(* IEC 61131-3 sources: plc-st-coding-agent/progress/evidence/f14_v11_public_20261113/jobs/custom_deepseek-v4pro, 104 files *)

(* ---- public-easy-01.candidate_01.st ---- *)
(* ENGINEERING_CONTRACT
Outputs by state (state is persistent across scans):
- Pump_Motor: ON in CLEANING; starts when bottleSensor TRUE from IDLE; OFF on cleaningConfirmButton. Retained while CLEANING, even if bottleSensor falls (PUB001/PUB002).
- Filling_Valve: ON in FILLING; starts on cleaningConfirmButton in CLEANING; OFF on fillingConfirmButton (PUB002/PUB003).
- Capping_Machine: ON in CAPPING; starts on fillingConfirmButton in FILLING; OFF on cappingConfirmButton (PUB003/PUB004).
- Packing_Machine: ON in PACKING; starts on cappingConfirmButton in CAPPING; OFF on packingConfirmButton (PUB004/PUB005).
- Completion_Light: ON in COMPLETE; starts on packingConfirmButton in PACKING; reset by finishedButton (PUB005/PUB006/PUB007).
Same-scan priority: one state transition per call via ELSIF chain; outputs are assigned after transition using final state.
Buttons are treated as level-sensitive; pulse width/protocol unspecified.
*)
(* CONTRACT_RULES [] *)

FUNCTION_BLOCK FillingLineControl
VAR_INPUT
    bottleSensor: BOOL;
    cleaningConfirmButton: BOOL;
    fillingConfirmButton: BOOL;
    cappingConfirmButton: BOOL;
    packingConfirmButton: BOOL;
    finishedButton: BOOL;
END_VAR
VAR_OUTPUT
    Pump_Motor: BOOL;
    Filling_Valve: BOOL;
    Capping_Machine: BOOL;
    Packing_Machine: BOOL;
    Completion_Light: BOOL;
END_VAR
VAR
    step: INT := 0; (* 0=IDLE, 1=CLEANING, 2=FILLING, 3=CAPPING, 4=PACKING, 5=COMPLETE *)
END_VAR

(* State transitions: at most one per scan *)
IF step = 0 THEN
    IF bottleSensor THEN
        step := 1;
    END_IF;
ELSIF step = 1 THEN
    IF cleaningConfirmButton THEN
        step := 2;
    END_IF;
ELSIF step = 2 THEN
    IF fillingConfirmButton THEN
        step := 3;
    END_IF;
ELSIF step = 3 THEN
    IF cappingConfirmButton THEN
        step := 4;
    END_IF;
ELSIF step = 4 THEN
    IF packingConfirmButton THEN
        step := 5;
    END_IF;
ELSIF step = 5 THEN
    IF finishedButton THEN
        step := 0;
    END_IF;
END_IF;

(* Output mapping based on final state *)
CASE step OF
    0:
        Pump_Motor := FALSE;
        Filling_Valve := FALSE;
        Capping_Machine := FALSE;
        Packing_Machine := FALSE;
        Completion_Light := FALSE;

    1:
        Pump_Motor := TRUE;
        Filling_Valve := FALSE;
        Capping_Machine := FALSE;
        Packing_Machine := FALSE;
        Completion_Light := FALSE;

    2:
        Pump_Motor := FALSE;
        Filling_Valve := TRUE;
        Capping_Machine := FALSE;
        Packing_Machine := FALSE;
        Completion_Light := FALSE;

    3:
        Pump_Motor := FALSE;
        Filling_Valve := FALSE;
        Capping_Machine := TRUE;
        Packing_Machine := FALSE;
        Completion_Light := FALSE;

    4:
        Pump_Motor := FALSE;
        Filling_Valve := FALSE;
        Capping_Machine := FALSE;
        Packing_Machine := TRUE;
        Completion_Light := FALSE;

    5:
        Pump_Motor := FALSE;
        Filling_Valve := FALSE;
        Capping_Machine := FALSE;
        Packing_Machine := FALSE;
        Completion_Light := TRUE;

    ELSE
        Pump_Motor := FALSE;
        Filling_Valve := FALSE;
        Capping_Machine := FALSE;
        Packing_Machine := FALSE;
        Completion_Light := FALSE;
END_CASE;

(* ---- public-easy-01.candidate_02.st ---- *)
(* ENGINEERING_CONTRACT
Outputs by state (state is persistent across scans):
- Pump_Motor: ON in CLEANING; starts when bottleSensor TRUE from IDLE; OFF on cleaningConfirmButton. Retained while CLEANING, even if bottleSensor falls (PUB001/PUB002).
- Filling_Valve: ON in FILLING; starts on cleaningConfirmButton in CLEANING; OFF on fillingConfirmButton (PUB002/PUB003).
- Capping_Machine: ON in CAPPING; starts on fillingConfirmButton in FILLING; OFF on cappingConfirmButton (PUB003/PUB004).
- Packing_Machine: ON in PACKING; starts on cappingConfirmButton in CAPPING; OFF on packingConfirmButton (PUB004/PUB005).
- Completion_Light: ON in COMPLETE; starts on packingConfirmButton in PACKING; reset by finishedButton (PUB005/PUB006/PUB007).
Same-scan priority: one state transition per call via ELSIF chain; outputs are assigned after transition using final state.
Buttons are treated as level-sensitive; pulse width/protocol unspecified.
*)
(* CONTRACT_RULES [] *)

FUNCTION_BLOCK FillingLineControl
VAR_INPUT
    bottleSensor: BOOL;
    cleaningConfirmButton: BOOL;
    fillingConfirmButton: BOOL;
    cappingConfirmButton: BOOL;
    packingConfirmButton: BOOL;
    finishedButton: BOOL;
END_VAR
VAR_OUTPUT
    Pump_Motor: BOOL;
    Filling_Valve: BOOL;
    Capping_Machine: BOOL;
    Packing_Machine: BOOL;
    Completion_Light: BOOL;
END_VAR
VAR
    step: INT := 0; (* 0=IDLE, 1=CLEANING, 2=FILLING, 3=CAPPING, 4=PACKING, 5=COMPLETE *)
END_VAR

(* State transitions: at most one per scan *)
IF step = 0 THEN
    IF bottleSensor THEN
        step := 1;
    END_IF;
ELSIF step = 1 THEN
    IF cleaningConfirmButton THEN
        step := 2;
    END_IF;
ELSIF step = 2 THEN
    IF fillingConfirmButton THEN
        step := 3;
    END_IF;
ELSIF step = 3 THEN
    IF cappingConfirmButton THEN
        step := 4;
    END_IF;
ELSIF step = 4 THEN
    IF packingConfirmButton THEN
        step := 5;
    END_IF;
ELSIF step = 5 THEN
    IF finishedButton THEN
        step := 0;
    END_IF;
END_IF;

(* Output mapping based on final state *)
CASE step OF
    0:
        Pump_Motor := FALSE;
        Filling_Valve := FALSE;
        Capping_Machine := FALSE;
        Packing_Machine := FALSE;
        Completion_Light := FALSE;

    1:
        Pump_Motor := TRUE;
        Filling_Valve := FALSE;
        Capping_Machine := FALSE;
        Packing_Machine := FALSE;
        Completion_Light := FALSE;

    2:
        Pump_Motor := FALSE;
        Filling_Valve := TRUE;
        Capping_Machine := FALSE;
        Packing_Machine := FALSE;
        Completion_Light := FALSE;

    3:
        Pump_Motor := FALSE;
        Filling_Valve := FALSE;
        Capping_Machine := TRUE;
        Packing_Machine := FALSE;
        Completion_Light := FALSE;

    4:
        Pump_Motor := FALSE;
        Filling_Valve := FALSE;
        Capping_Machine := FALSE;
        Packing_Machine := TRUE;
        Completion_Light := FALSE;

    5:
        Pump_Motor := FALSE;
        Filling_Valve := FALSE;
        Capping_Machine := FALSE;
        Packing_Machine := FALSE;
        Completion_Light := TRUE;

    ELSE
        Pump_Motor := FALSE;
        Filling_Valve := FALSE;
        Capping_Machine := FALSE;
        Packing_Machine := FALSE;
        Completion_Light := FALSE;
END_CASE;

END_FUNCTION_BLOCK

(* ---- public-easy-01.candidate_03.st ---- *)
(* ENGINEERING_CONTRACT
Outputs by state (state is persistent across scans):
- Pump_Motor: ON in CLEANING; starts when bottleSensor TRUE from IDLE; OFF on cleaningConfirmButton. Retained while CLEANING, even if bottleSensor falls (PUB001/PUB002).
- Filling_Valve: ON in FILLING; starts on cleaningConfirmButton in CLEANING; OFF on fillingConfirmButton (PUB002/PUB003).
- Capping_Machine: ON in CAPPING; starts on fillingConfirmButton in FILLING; OFF on cappingConfirmButton (PUB003/PUB004).
- Packing_Machine: ON in PACKING; starts on cappingConfirmButton in CAPPING; OFF on packingConfirmButton (PUB004/PUB005).
- Completion_Light: ON in COMPLETE; starts on packingConfirmButton in PACKING; reset by finishedButton (PUB005/PUB006/PUB007).
Same-scan priority:
- Primary ELSIF chain processes one normal step.
- If finishedButton resets to IDLE and bottleSensor is already TRUE, re-enter CLEANING immediately in same scan.
Outputs are assigned after transition logic using final state.
Buttons are treated as level-sensitive; pulse width/protocol unspecified.
*)
(* CONTRACT_RULES [] *)

FUNCTION_BLOCK FillingLineControl
VAR_INPUT
    bottleSensor: BOOL;
    cleaningConfirmButton: BOOL;
    fillingConfirmButton: BOOL;
    cappingConfirmButton: BOOL;
    packingConfirmButton: BOOL;
    finishedButton: BOOL;
END_VAR
VAR_OUTPUT
    Pump_Motor: BOOL;
    Filling_Valve: BOOL;
    Capping_Machine: BOOL;
    Packing_Machine: BOOL;
    Completion_Light: BOOL;
END_VAR
VAR
    step: INT := 0; (* 0=IDLE, 1=CLEANING, 2=FILLING, 3=CAPPING, 4=PACKING, 5=COMPLETE *)
END_VAR

(* Primary state transitions: at most one normal step per scan *)
IF step = 0 THEN
    IF bottleSensor THEN
        step := 1;
    END_IF;
ELSIF step = 1 THEN
    IF cleaningConfirmButton THEN
        step := 2;
    END_IF;
ELSIF step = 2 THEN
    IF fillingConfirmButton THEN
        step := 3;
    END_IF;
ELSIF step = 3 THEN
    IF cappingConfirmButton THEN
        step := 4;
    END_IF;
ELSIF step = 4 THEN
    IF packingConfirmButton THEN
        step := 5;
    END_IF;
ELSIF step = 5 THEN
    IF finishedButton THEN
        step := 0;
    END_IF;
END_IF;

(* Same-scan reactivation: if finished just reset state to IDLE and a bottle is
   already detected, start cleaning immediately instead of waiting one scan. *)
IF step = 0 THEN
    IF bottleSensor THEN
        step := 1;
    END_IF;
END_IF;

(* Output mapping based on final state *)
CASE step OF
    0:
        Pump_Motor := FALSE;
        Filling_Valve := FALSE;
        Capping_Machine := FALSE;
        Packing_Machine := FALSE;
        Completion_Light := FALSE;

    1:
        Pump_Motor := TRUE;
        Filling_Valve := FALSE;
        Capping_Machine := FALSE;
        Packing_Machine := FALSE;
        Completion_Light := FALSE;

    2:
        Pump_Motor := FALSE;
        Filling_Valve := TRUE;
        Capping_Machine := FALSE;
        Packing_Machine := FALSE;
        Completion_Light := FALSE;

    3:
        Pump_Motor := FALSE;
        Filling_Valve := FALSE;
        Capping_Machine := TRUE;
        Packing_Machine := FALSE;
        Completion_Light := FALSE;

    4:
        Pump_Motor := FALSE;
        Filling_Valve := FALSE;
        Capping_Machine := FALSE;
        Packing_Machine := TRUE;
        Completion_Light := FALSE;

    5:
        Pump_Motor := FALSE;
        Filling_Valve := FALSE;
        Capping_Machine := FALSE;
        Packing_Machine := FALSE;
        Completion_Light := TRUE;

    ELSE
        Pump_Motor := FALSE;
        Filling_Valve := FALSE;
        Capping_Machine := FALSE;
        Packing_Machine := FALSE;
        Completion_Light := FALSE;
END_CASE;

END_FUNCTION_BLOCK

(* ---- public-easy-01.candidate_04.st ---- *)
(* ENGINEERING_CONTRACT
Outputs by state (state is persistent across scans):
- Pump_Motor: ON in CLEANING; starts when bottleSensor TRUE from IDLE; OFF on cleaningConfirmButton. Retained while CLEANING, even if bottleSensor falls (PUB001/PUB002).
- Filling_Valve: ON in FILLING; starts on cleaningConfirmButton in CLEANING; OFF on fillingConfirmButton (PUB002/PUB003).
- Capping_Machine: ON in CAPPING; starts on fillingConfirmButton in FILLING; OFF on cappingConfirmButton (PUB003/PUB004).
- Packing_Machine: ON in PACKING; starts on cappingConfirmButton in CAPPING; OFF on packingConfirmButton (PUB004/PUB005).
- Completion_Light: ON in COMPLETE; starts on packingConfirmButton in PACKING; reset by finishedButton (PUB005/PUB006/PUB007).
Same-scan priority:
- Primary ELSIF chain processes one normal step.
- If finishedButton resets to IDLE and bottleSensor is already TRUE, re-enter CLEANING immediately in same scan.
Outputs are assigned after transition logic using final state.
Buttons are treated as level-sensitive; pulse width/protocol unspecified.
*)
(* CONTRACT_RULES [
  {"kind":"hold_until_reset","output":"Pump_Motor","set_input":"bottleSensor","reset_input":"cleaningConfirmButton"},
  {"kind":"hold_until_reset","output":"Filling_Valve","set_input":"cleaningConfirmButton","reset_input":"fillingConfirmButton"},
  {"kind":"hold_until_reset","output":"Capping_Machine","set_input":"fillingConfirmButton","reset_input":"cappingConfirmButton"},
  {"kind":"hold_until_reset","output":"Packing_Machine","set_input":"cappingConfirmButton","reset_input":"packingConfirmButton"},
  {"kind":"hold_until_reset","output":"Completion_Light","set_input":"packingConfirmButton","reset_input":"finishedButton"}
] *)

FUNCTION_BLOCK FillingLineControl
VAR_INPUT
    bottleSensor: BOOL;
    cleaningConfirmButton: BOOL;
    fillingConfirmButton: BOOL;
    cappingConfirmButton: BOOL;
    packingConfirmButton: BOOL;
    finishedButton: BOOL;
END_VAR
VAR_OUTPUT
    Pump_Motor: BOOL;
    Filling_Valve: BOOL;
    Capping_Machine: BOOL;
    Packing_Machine: BOOL;
    Completion_Light: BOOL;
END_VAR
VAR
    step: INT := 0; (* 0=IDLE, 1=CLEANING, 2=FILLING, 3=CAPPING, 4=PACKING, 5=COMPLETE *)
END_VAR

(* Primary state transitions: at most one normal step per scan *)
IF step = 0 THEN
    IF bottleSensor THEN
        step := 1;
    END_IF;
ELSIF step = 1 THEN
    IF cleaningConfirmButton THEN
        step := 2;
    END_IF;
ELSIF step = 2 THEN
    IF fillingConfirmButton THEN
        step := 3;
    END_IF;
ELSIF step = 3 THEN
    IF cappingConfirmButton THEN
        step := 4;
    END_IF;
ELSIF step = 4 THEN
    IF packingConfirmButton THEN
        step := 5;
    END_IF;
ELSIF step = 5 THEN
    IF finishedButton THEN
        step := 0;
    END_IF;
END_IF;

(* Same-scan reactivation: if finished just reset state to IDLE and a bottle is
   already detected, start cleaning immediately instead of waiting one scan. *)
IF step = 0 THEN
    IF bottleSensor THEN
        step := 1;
    END_IF;
END_IF;

(* Output mapping based on final state *)
CASE step OF
    0:
        Pump_Motor := FALSE;
        Filling_Valve := FALSE;
        Capping_Machine := FALSE;
        Packing_Machine := FALSE;
        Completion_Light := FALSE;

    1:
        Pump_Motor := TRUE;
        Filling_Valve := FALSE;
        Capping_Machine := FALSE;
        Packing_Machine := FALSE;
        Completion_Light := FALSE;

    2:
        Pump_Motor := FALSE;
        Filling_Valve := TRUE;
        Capping_Machine := FALSE;
        Packing_Machine := FALSE;
        Completion_Light := FALSE;

    3:
        Pump_Motor := FALSE;
        Filling_Valve := FALSE;
        Capping_Machine := TRUE;
        Packing_Machine := FALSE;
        Completion_Light := FALSE;

    4:
        Pump_Motor := FALSE;
        Filling_Valve := FALSE;
        Capping_Machine := FALSE;
        Packing_Machine := TRUE;
        Completion_Light := FALSE;

    5:
        Pump_Motor := FALSE;
        Filling_Valve := FALSE;
        Capping_Machine := FALSE;
        Packing_Machine := FALSE;
        Completion_Light := TRUE;

    ELSE
        Pump_Motor := FALSE;
        Filling_Valve := FALSE;
        Capping_Machine := FALSE;
        Packing_Machine := FALSE;
        Completion_Light := FALSE;
END_CASE;

END_FUNCTION_BLOCK

(* ---- public-easy-01.raw_candidate_01.st ---- *)
(* ENGINEERING_CONTRACT
Outputs by state (state is persistent across scans):
- Pump_Motor: ON in CLEANING; starts when bottleSensor TRUE from IDLE; OFF on cleaningConfirmButton. Retained while CLEANING, even if bottleSensor falls (PUB001/PUB002).
- Filling_Valve: ON in FILLING; starts on cleaningConfirmButton in CLEANING; OFF on fillingConfirmButton (PUB002/PUB003).
- Capping_Machine: ON in CAPPING; starts on fillingConfirmButton in FILLING; OFF on cappingConfirmButton (PUB003/PUB004).
- Packing_Machine: ON in PACKING; starts on cappingConfirmButton in CAPPING; OFF on packingConfirmButton (PUB004/PUB005).
- Completion_Light: ON in COMPLETE; starts on packingConfirmButton in PACKING; reset by finishedButton (PUB005/PUB006/PUB007).
Same-scan priority: one state transition per call via ELSIF chain; outputs are assigned after transition using final state.
Buttons are treated as level-sensitive; pulse width/protocol unspecified.
*)
(* CONTRACT_RULES [] *)

FUNCTION_BLOCK FillingLineControl
VAR_INPUT
    bottleSensor: BOOL;
    cleaningConfirmButton: BOOL;
    fillingConfirmButton: BOOL;
    cappingConfirmButton: BOOL;
    packingConfirmButton: BOOL;
    finishedButton: BOOL;
END_VAR
VAR_OUTPUT
    Pump_Motor: BOOL;
    Filling_Valve: BOOL;
    Capping_Machine: BOOL;
    Packing_Machine: BOOL;
    Completion_Light: BOOL;
END_VAR
VAR
    step: INT := 0; (* 0=IDLE, 1=CLEANING, 2=FILLING, 3=CAPPING, 4=PACKING, 5=COMPLETE *)
END_VAR

(* State transitions: at most one per scan *)
IF step = 0 THEN
    IF bottleSensor THEN
        step := 1;
    END_IF;
ELSIF step = 1 THEN
    IF cleaningConfirmButton THEN
        step := 2;
    END_IF;
ELSIF step = 2 THEN
    IF fillingConfirmButton THEN
        step := 3;
    END_IF;
ELSIF step = 3 THEN
    IF cappingConfirmButton THEN
        step := 4;
    END_IF;
ELSIF step = 4 THEN
    IF packingConfirmButton THEN
        step := 5;
    END_IF;
ELSIF step = 5 THEN
    IF finishedButton THEN
        step := 0;
    END_IF;
END_IF;

(* Output mapping based on final state *)
CASE step OF
    0:
        Pump_Motor := FALSE;
        Filling_Valve := FALSE;
        Capping_Machine := FALSE;
        Packing_Machine := FALSE;
        Completion_Light := FALSE;

    1:
        Pump_Motor := TRUE;
        Filling_Valve := FALSE;
        Capping_Machine := FALSE;
        Packing_Machine := FALSE;
        Completion_Light := FALSE;

    2:
        Pump_Motor := FALSE;
        Filling_Valve := TRUE;
        Capping_Machine := FALSE;
        Packing_Machine := FALSE;
        Completion_Light := FALSE;

    3:
        Pump_Motor := FALSE;
        Filling_Valve := FALSE;
        Capping_Machine := TRUE;
        Packing_Machine := FALSE;
        Completion_Light := FALSE;

    4:
        Pump_Motor := FALSE;
        Filling_Valve := FALSE;
        Capping_Machine := FALSE;
        Packing_Machine := TRUE;
        Completion_Light := FALSE;

    5:
        Pump_Motor := FALSE;
        Filling_Valve := FALSE;
        Capping_Machine := FALSE;
        Packing_Machine := FALSE;
        Completion_Light := TRUE;

    ELSE
        Pump_Motor := FALSE;
        Filling_Valve := FALSE;
        Capping_Machine := FALSE;
        Packing_Machine := FALSE;
        Completion_Light := FALSE;
END_CASE;

(* ---- public-easy-01.raw_candidate_02.st ---- *)
(* ENGINEERING_CONTRACT
Outputs by state (state is persistent across scans):
- Pump_Motor: ON in CLEANING; starts when bottleSensor TRUE from IDLE; OFF on cleaningConfirmButton. Retained while CLEANING, even if bottleSensor falls (PUB001/PUB002).
- Filling_Valve: ON in FILLING; starts on cleaningConfirmButton in CLEANING; OFF on fillingConfirmButton (PUB002/PUB003).
- Capping_Machine: ON in CAPPING; starts on fillingConfirmButton in FILLING; OFF on cappingConfirmButton (PUB003/PUB004).
- Packing_Machine: ON in PACKING; starts on cappingConfirmButton in CAPPING; OFF on packingConfirmButton (PUB004/PUB005).
- Completion_Light: ON in COMPLETE; starts on packingConfirmButton in PACKING; reset by finishedButton (PUB005/PUB006/PUB007).
Same-scan priority: one state transition per call via ELSIF chain; outputs are assigned after transition using final state.
Buttons are treated as level-sensitive; pulse width/protocol unspecified.
*)
(* CONTRACT_RULES [] *)

FUNCTION_BLOCK FillingLineControl
VAR_INPUT
    bottleSensor: BOOL;
    cleaningConfirmButton: BOOL;
    fillingConfirmButton: BOOL;
    cappingConfirmButton: BOOL;
    packingConfirmButton: BOOL;
    finishedButton: BOOL;
END_VAR
VAR_OUTPUT
    Pump_Motor: BOOL;
    Filling_Valve: BOOL;
    Capping_Machine: BOOL;
    Packing_Machine: BOOL;
    Completion_Light: BOOL;
END_VAR
VAR
    step: INT := 0; (* 0=IDLE, 1=CLEANING, 2=FILLING, 3=CAPPING, 4=PACKING, 5=COMPLETE *)
END_VAR

(* State transitions: at most one per scan *)
IF step = 0 THEN
    IF bottleSensor THEN
        step := 1;
    END_IF;
ELSIF step = 1 THEN
    IF cleaningConfirmButton THEN
        step := 2;
    END_IF;
ELSIF step = 2 THEN
    IF fillingConfirmButton THEN
        step := 3;
    END_IF;
ELSIF step = 3 THEN
    IF cappingConfirmButton THEN
        step := 4;
    END_IF;
ELSIF step = 4 THEN
    IF packingConfirmButton THEN
        step := 5;
    END_IF;
ELSIF step = 5 THEN
    IF finishedButton THEN
        step := 0;
    END_IF;
END_IF;

(* Output mapping based on final state *)
CASE step OF
    0:
        Pump_Motor := FALSE;
        Filling_Valve := FALSE;
        Capping_Machine := FALSE;
        Packing_Machine := FALSE;
        Completion_Light := FALSE;

    1:
        Pump_Motor := TRUE;
        Filling_Valve := FALSE;
        Capping_Machine := FALSE;
        Packing_Machine := FALSE;
        Completion_Light := FALSE;

    2:
        Pump_Motor := FALSE;
        Filling_Valve := TRUE;
        Capping_Machine := FALSE;
        Packing_Machine := FALSE;
        Completion_Light := FALSE;

    3:
        Pump_Motor := FALSE;
        Filling_Valve := FALSE;
        Capping_Machine := TRUE;
        Packing_Machine := FALSE;
        Completion_Light := FALSE;

    4:
        Pump_Motor := FALSE;
        Filling_Valve := FALSE;
        Capping_Machine := FALSE;
        Packing_Machine := TRUE;
        Completion_Light := FALSE;

    5:
        Pump_Motor := FALSE;
        Filling_Valve := FALSE;
        Capping_Machine := FALSE;
        Packing_Machine := FALSE;
        Completion_Light := TRUE;

    ELSE
        Pump_Motor := FALSE;
        Filling_Valve := FALSE;
        Capping_Machine := FALSE;
        Packing_Machine := FALSE;
        Completion_Light := FALSE;
END_CASE;

END_FUNCTION_BLOCK

(* ---- public-easy-01.raw_candidate_03.st ---- *)
(* ENGINEERING_CONTRACT
Outputs by state (state is persistent across scans):
- Pump_Motor: ON in CLEANING; starts when bottleSensor TRUE from IDLE; OFF on cleaningConfirmButton. Retained while CLEANING, even if bottleSensor falls (PUB001/PUB002).
- Filling_Valve: ON in FILLING; starts on cleaningConfirmButton in CLEANING; OFF on fillingConfirmButton (PUB002/PUB003).
- Capping_Machine: ON in CAPPING; starts on fillingConfirmButton in FILLING; OFF on cappingConfirmButton (PUB003/PUB004).
- Packing_Machine: ON in PACKING; starts on cappingConfirmButton in CAPPING; OFF on packingConfirmButton (PUB004/PUB005).
- Completion_Light: ON in COMPLETE; starts on packingConfirmButton in PACKING; reset by finishedButton (PUB005/PUB006/PUB007).
Same-scan priority:
- Primary ELSIF chain processes one normal step.
- If finishedButton resets to IDLE and bottleSensor is already TRUE, re-enter CLEANING immediately in same scan.
Outputs are assigned after transition logic using final state.
Buttons are treated as level-sensitive; pulse width/protocol unspecified.
*)
(* CONTRACT_RULES [] *)

FUNCTION_BLOCK FillingLineControl
VAR_INPUT
    bottleSensor: BOOL;
    cleaningConfirmButton: BOOL;
    fillingConfirmButton: BOOL;
    cappingConfirmButton: BOOL;
    packingConfirmButton: BOOL;
    finishedButton: BOOL;
END_VAR
VAR_OUTPUT
    Pump_Motor: BOOL;
    Filling_Valve: BOOL;
    Capping_Machine: BOOL;
    Packing_Machine: BOOL;
    Completion_Light: BOOL;
END_VAR
VAR
    step: INT := 0; (* 0=IDLE, 1=CLEANING, 2=FILLING, 3=CAPPING, 4=PACKING, 5=COMPLETE *)
END_VAR

(* Primary state transitions: at most one normal step per scan *)
IF step = 0 THEN
    IF bottleSensor THEN
        step := 1;
    END_IF;
ELSIF step = 1 THEN
    IF cleaningConfirmButton THEN
        step := 2;
    END_IF;
ELSIF step = 2 THEN
    IF fillingConfirmButton THEN
        step := 3;
    END_IF;
ELSIF step = 3 THEN
    IF cappingConfirmButton THEN
        step := 4;
    END_IF;
ELSIF step = 4 THEN
    IF packingConfirmButton THEN
        step := 5;
    END_IF;
ELSIF step = 5 THEN
    IF finishedButton THEN
        step := 0;
    END_IF;
END_IF;

(* Same-scan reactivation: if finished just reset state to IDLE and a bottle is
   already detected, start cleaning immediately instead of waiting one scan. *)
IF step = 0 THEN
    IF bottleSensor THEN
        step := 1;
    END_IF;
END_IF;

(* Output mapping based on final state *)
CASE step OF
    0:
        Pump_Motor := FALSE;
        Filling_Valve := FALSE;
        Capping_Machine := FALSE;
        Packing_Machine := FALSE;
        Completion_Light := FALSE;

    1:
        Pump_Motor := TRUE;
        Filling_Valve := FALSE;
        Capping_Machine := FALSE;
        Packing_Machine := FALSE;
        Completion_Light := FALSE;

    2:
        Pump_Motor := FALSE;
        Filling_Valve := TRUE;
        Capping_Machine := FALSE;
        Packing_Machine := FALSE;
        Completion_Light := FALSE;

    3:
        Pump_Motor := FALSE;
        Filling_Valve := FALSE;
        Capping_Machine := TRUE;
        Packing_Machine := FALSE;
        Completion_Light := FALSE;

    4:
        Pump_Motor := FALSE;
        Filling_Valve := FALSE;
        Capping_Machine := FALSE;
        Packing_Machine := TRUE;
        Completion_Light := FALSE;

    5:
        Pump_Motor := FALSE;
        Filling_Valve := FALSE;
        Capping_Machine := FALSE;
        Packing_Machine := FALSE;
        Completion_Light := TRUE;

    ELSE
        Pump_Motor := FALSE;
        Filling_Valve := FALSE;
        Capping_Machine := FALSE;
        Packing_Machine := FALSE;
        Completion_Light := FALSE;
END_CASE;

END_FUNCTION_BLOCK

(* ---- public-easy-01.raw_candidate_04.st ---- *)
(* ENGINEERING_CONTRACT
Outputs by state (state is persistent across scans):
- Pump_Motor: ON in CLEANING; starts when bottleSensor TRUE from IDLE; OFF on cleaningConfirmButton. Retained while CLEANING, even if bottleSensor falls (PUB001/PUB002).
- Filling_Valve: ON in FILLING; starts on cleaningConfirmButton in CLEANING; OFF on fillingConfirmButton (PUB002/PUB003).
- Capping_Machine: ON in CAPPING; starts on fillingConfirmButton in FILLING; OFF on cappingConfirmButton (PUB003/PUB004).
- Packing_Machine: ON in PACKING; starts on cappingConfirmButton in CAPPING; OFF on packingConfirmButton (PUB004/PUB005).
- Completion_Light: ON in COMPLETE; starts on packingConfirmButton in PACKING; reset by finishedButton (PUB005/PUB006/PUB007).
Same-scan priority:
- Primary ELSIF chain processes one normal step.
- If finishedButton resets to IDLE and bottleSensor is already TRUE, re-enter CLEANING immediately in same scan.
Outputs are assigned after transition logic using final state.
Buttons are treated as level-sensitive; pulse width/protocol unspecified.
*)
(* CONTRACT_RULES [
  {"kind":"hold_until_reset","output":"Pump_Motor","set_input":"bottleSensor","reset_input":"cleaningConfirmButton"},
  {"kind":"hold_until_reset","output":"Filling_Valve","set_input":"cleaningConfirmButton","reset_input":"fillingConfirmButton"},
  {"kind":"hold_until_reset","output":"Capping_Machine","set_input":"fillingConfirmButton","reset_input":"cappingConfirmButton"},
  {"kind":"hold_until_reset","output":"Packing_Machine","set_input":"cappingConfirmButton","reset_input":"packingConfirmButton"},
  {"kind":"hold_until_reset","output":"Completion_Light","set_input":"packingConfirmButton","reset_input":"finishedButton"}
] *)

FUNCTION_BLOCK FillingLineControl
VAR_INPUT
    bottleSensor: BOOL;
    cleaningConfirmButton: BOOL;
    fillingConfirmButton: BOOL;
    cappingConfirmButton: BOOL;
    packingConfirmButton: BOOL;
    finishedButton: BOOL;
END_VAR
VAR_OUTPUT
    Pump_Motor: BOOL;
    Filling_Valve: BOOL;
    Capping_Machine: BOOL;
    Packing_Machine: BOOL;
    Completion_Light: BOOL;
END_VAR
VAR
    step: INT := 0; (* 0=IDLE, 1=CLEANING, 2=FILLING, 3=CAPPING, 4=PACKING, 5=COMPLETE *)
END_VAR

(* Primary state transitions: at most one normal step per scan *)
IF step = 0 THEN
    IF bottleSensor THEN
        step := 1;
    END_IF;
ELSIF step = 1 THEN
    IF cleaningConfirmButton THEN
        step := 2;
    END_IF;
ELSIF step = 2 THEN
    IF fillingConfirmButton THEN
        step := 3;
    END_IF;
ELSIF step = 3 THEN
    IF cappingConfirmButton THEN
        step := 4;
    END_IF;
ELSIF step = 4 THEN
    IF packingConfirmButton THEN
        step := 5;
    END_IF;
ELSIF step = 5 THEN
    IF finishedButton THEN
        step := 0;
    END_IF;
END_IF;

(* Same-scan reactivation: if finished just reset state to IDLE and a bottle is
   already detected, start cleaning immediately instead of waiting one scan. *)
IF step = 0 THEN
    IF bottleSensor THEN
        step := 1;
    END_IF;
END_IF;

(* Output mapping based on final state *)
CASE step OF
    0:
        Pump_Motor := FALSE;
        Filling_Valve := FALSE;
        Capping_Machine := FALSE;
        Packing_Machine := FALSE;
        Completion_Light := FALSE;

    1:
        Pump_Motor := TRUE;
        Filling_Valve := FALSE;
        Capping_Machine := FALSE;
        Packing_Machine := FALSE;
        Completion_Light := FALSE;

    2:
        Pump_Motor := FALSE;
        Filling_Valve := TRUE;
        Capping_Machine := FALSE;
        Packing_Machine := FALSE;
        Completion_Light := FALSE;

    3:
        Pump_Motor := FALSE;
        Filling_Valve := FALSE;
        Capping_Machine := TRUE;
        Packing_Machine := FALSE;
        Completion_Light := FALSE;

    4:
        Pump_Motor := FALSE;
        Filling_Valve := FALSE;
        Capping_Machine := FALSE;
        Packing_Machine := TRUE;
        Completion_Light := FALSE;

    5:
        Pump_Motor := FALSE;
        Filling_Valve := FALSE;
        Capping_Machine := FALSE;
        Packing_Machine := FALSE;
        Completion_Light := TRUE;

    ELSE
        Pump_Motor := FALSE;
        Filling_Valve := FALSE;
        Capping_Machine := FALSE;
        Packing_Machine := FALSE;
        Completion_Light := FALSE;
END_CASE;

END_FUNCTION_BLOCK

(* ---- public-easy-02.candidate_01.st ---- *)
FUNCTION_BLOCK FB
(* ENGINEERING_CONTRACT
   PUB001: every scan compares DWORD input value against the previous scan value.
   hasChanged: combinational this scan; TRUE iff current value <> stored previous value.
   hasRisingEdges/risingBits/noOfRisingBits: combinational this scan; rising mask = current AND NOT previous.
   hasFallingEdges/fallingBits/noOfFallingBits: combinational this scan; falling mask = previous AND NOT current.
   No output is latched; all edge outputs return to FALSE/0 on the next equal-value scan.
   First scan initializes previous value to current value, so no change or edge is reported at startup.
   Counts are USINT bit counts 0..32; masks are DWORD bit positions 0..31.
*)
(* CONTRACT_RULES [] *)
VAR_INPUT
    value : DWORD;
END_VAR
VAR_OUTPUT
    hasChanged : BOOL;
    hasRisingEdges : BOOL;
    risingBits : DWORD;
    noOfRisingBits : USINT;
    hasFallingEdges : BOOL;
    fallingBits : DWORD;
    noOfFallingBits : USINT;
END_VAR
VAR
    local_initialized : BOOL := FALSE;
    lastValue : DWORD;
    tmp_i : DINT;
    tmp_shift : UDINT;
    tmp_mask : DWORD;
END_VAR

IF NOT local_initialized THEN
    local_initialized := TRUE;
    lastValue := value;
    hasChanged := FALSE;
    hasRisingEdges := FALSE;
    risingBits := 0;
    noOfRisingBits := 0;
    hasFallingEdges := FALSE;
    fallingBits := 0;
    noOfFallingBits := 0;
    RETURN;
END_IF;

hasChanged := value <> lastValue;

IF hasChanged THEN
    risingBits := value AND (NOT lastValue);
    fallingBits := lastValue AND (NOT value);
    noOfRisingBits := 0;
    noOfFallingBits := 0;

    FOR tmp_i := 0 TO 31 DO
        tmp_shift := DINT_TO_UDINT(tmp_i);
        tmp_mask := SHL(DWORD#1, tmp_shift);

        IF (risingBits AND tmp_mask) <> DWORD#0 THEN
            noOfRisingBits := noOfRisingBits + 1;
        END_IF;

        IF (fallingBits AND tmp_mask) <> DWORD#0 THEN
            noOfFallingBits := noOfFallingBits + 1;
        END_IF;
    END_FOR;

    hasRisingEdges := noOfRisingBits > 0;
    hasFallingEdges := noOfFallingBits > 0;
ELSE
    hasRisingEdges := FALSE;
    risingBits := 0;
    noOfRisingBits := 0;
    hasFallingEdges := FALSE;
    fallingBits := 0;
    noOfFallingBits := 0;
END_IF;

lastValue := value;
END_FUNCTION_BLOCK

(* ---- public-easy-02.candidate_02.st ---- *)
FUNCTION_BLOCK FB
(* ENGINEERING_CONTRACT
   PUB001: every scan compares DWORD input value against stored previous value (initial 0).
   hasChanged: combinational this scan; TRUE iff current value <> stored previous value.
   hasRisingEdges/risingBits/noOfRisingBits: combinational this scan; rising mask = current AND NOT previous.
   hasFallingEdges/fallingBits/noOfFallingBits: combinational this scan; falling mask = previous AND NOT current.
   No output is latched; all edge outputs return to FALSE/0 on the next equal-value scan.
   First scan compares against default previous value 0, so edges from 0 are detected.
   Counts are USINT bit counts 0..32; masks are DWORD bit positions 0..31.
*)
(* CONTRACT_RULES [] *)
VAR_INPUT
    value : DWORD;
END_VAR
VAR_OUTPUT
    hasChanged : BOOL;
    hasRisingEdges : BOOL;
    risingBits : DWORD;
    noOfRisingBits : USINT;
    hasFallingEdges : BOOL;
    fallingBits : DWORD;
    noOfFallingBits : USINT;
END_VAR
VAR
    lastValue : DWORD; (* defaults to 0 *)
    tmp_i : DINT;
    tmp_shift : UDINT;
    tmp_mask : DWORD;
END_VAR

hasChanged := value <> lastValue;

IF hasChanged THEN
    risingBits := value AND (NOT lastValue);
    fallingBits := lastValue AND (NOT value);
    noOfRisingBits := 0;
    noOfFallingBits := 0;

    FOR tmp_i := 0 TO 31 DO
        tmp_shift := DINT_TO_UDINT(tmp_i);
        tmp_mask := SHL(DWORD#1, tmp_shift);

        IF (risingBits AND tmp_mask) <> DWORD#0 THEN
            noOfRisingBits := noOfRisingBits + 1;
        END_IF;

        IF (fallingBits AND tmp_mask) <> DWORD#0 THEN
            noOfFallingBits := noOfFallingBits + 1;
        END_IF;
    END_FOR;

    hasRisingEdges := noOfRisingBits > 0;
    hasFallingEdges := noOfFallingBits > 0;
ELSE
    hasRisingEdges := FALSE;
    risingBits := 0;
    noOfRisingBits := 0;
    hasFallingEdges := FALSE;
    fallingBits := 0;
    noOfFallingBits := 0;
END_IF;

lastValue := value;
END_FUNCTION_BLOCK

(* ---- public-easy-02.raw_candidate_01.st ---- *)
FUNCTION_BLOCK FB
(* ENGINEERING_CONTRACT
   PUB001: every scan compares DWORD input value against the previous scan value.
   hasChanged: combinational this scan; TRUE iff current value <> stored previous value.
   hasRisingEdges/risingBits/noOfRisingBits: combinational this scan; rising mask = current AND NOT previous.
   hasFallingEdges/fallingBits/noOfFallingBits: combinational this scan; falling mask = previous AND NOT current.
   No output is latched; all edge outputs return to FALSE/0 on the next equal-value scan.
   First scan initializes previous value to current value, so no change or edge is reported at startup.
   Counts are USINT bit counts 0..32; masks are DWORD bit positions 0..31.
*)
(* CONTRACT_RULES [] *)
VAR_INPUT
    value : DWORD;
END_VAR
VAR_OUTPUT
    hasChanged : BOOL;
    hasRisingEdges : BOOL;
    risingBits : DWORD;
    noOfRisingBits : USINT;
    hasFallingEdges : BOOL;
    fallingBits : DWORD;
    noOfFallingBits : USINT;
END_VAR
VAR
    local_initialized : BOOL := FALSE;
    lastValue : DWORD;
    tmp_i : DINT;
    tmp_shift : UDINT;
    tmp_mask : DWORD;
END_VAR

IF NOT local_initialized THEN
    local_initialized := TRUE;
    lastValue := value;
    hasChanged := FALSE;
    hasRisingEdges := FALSE;
    risingBits := 0;
    noOfRisingBits := 0;
    hasFallingEdges := FALSE;
    fallingBits := 0;
    noOfFallingBits := 0;
    RETURN;
END_IF;

hasChanged := value <> lastValue;

IF hasChanged THEN
    risingBits := value AND (NOT lastValue);
    fallingBits := lastValue AND (NOT value);
    noOfRisingBits := 0;
    noOfFallingBits := 0;

    FOR tmp_i := 0 TO 31 DO
        tmp_shift := DINT_TO_UDINT(tmp_i);
        tmp_mask := SHL(DWORD#1, tmp_shift);

        IF (risingBits AND tmp_mask) <> DWORD#0 THEN
            noOfRisingBits := noOfRisingBits + 1;
        END_IF;

        IF (fallingBits AND tmp_mask) <> DWORD#0 THEN
            noOfFallingBits := noOfFallingBits + 1;
        END_IF;
    END_FOR;

    hasRisingEdges := noOfRisingBits > 0;
    hasFallingEdges := noOfFallingBits > 0;
ELSE
    hasRisingEdges := FALSE;
    risingBits := 0;
    noOfRisingBits := 0;
    hasFallingEdges := FALSE;
    fallingBits := 0;
    noOfFallingBits := 0;
END_IF;

lastValue := value;
END_FUNCTION_BLOCK

(* ---- public-easy-02.raw_candidate_02.st ---- *)
FUNCTION_BLOCK FB
(* ENGINEERING_CONTRACT
   PUB001: every scan compares DWORD input value against stored previous value (initial 0).
   hasChanged: combinational this scan; TRUE iff current value <> stored previous value.
   hasRisingEdges/risingBits/noOfRisingBits: combinational this scan; rising mask = current AND NOT previous.
   hasFallingEdges/fallingBits/noOfFallingBits: combinational this scan; falling mask = previous AND NOT current.
   No output is latched; all edge outputs return to FALSE/0 on the next equal-value scan.
   First scan compares against default previous value 0, so edges from 0 are detected.
   Counts are USINT bit counts 0..32; masks are DWORD bit positions 0..31.
*)
(* CONTRACT_RULES [] *)
VAR_INPUT
    value : DWORD;
END_VAR
VAR_OUTPUT
    hasChanged : BOOL;
    hasRisingEdges : BOOL;
    risingBits : DWORD;
    noOfRisingBits : USINT;
    hasFallingEdges : BOOL;
    fallingBits : DWORD;
    noOfFallingBits : USINT;
END_VAR
VAR
    lastValue : DWORD; (* defaults to 0 *)
    tmp_i : DINT;
    tmp_shift : UDINT;
    tmp_mask : DWORD;
END_VAR

hasChanged := value <> lastValue;

IF hasChanged THEN
    risingBits := value AND (NOT lastValue);
    fallingBits := lastValue AND (NOT value);
    noOfRisingBits := 0;
    noOfFallingBits := 0;

    FOR tmp_i := 0 TO 31 DO
        tmp_shift := DINT_TO_UDINT(tmp_i);
        tmp_mask := SHL(DWORD#1, tmp_shift);

        IF (risingBits AND tmp_mask) <> DWORD#0 THEN
            noOfRisingBits := noOfRisingBits + 1;
        END_IF;

        IF (fallingBits AND tmp_mask) <> DWORD#0 THEN
            noOfFallingBits := noOfFallingBits + 1;
        END_IF;
    END_FOR;

    hasRisingEdges := noOfRisingBits > 0;
    hasFallingEdges := noOfFallingBits > 0;
ELSE
    hasRisingEdges := FALSE;
    risingBits := 0;
    noOfRisingBits := 0;
    hasFallingEdges := FALSE;
    fallingBits := 0;
    noOfFallingBits := 0;
END_IF;

lastValue := value;
END_FUNCTION_BLOCK

(* ---- public-easy-03.candidate_01.st ---- *)
FUNCTION_BLOCK AlarmHandling
VAR_INPUT
    Value : REAL;
    hiLevel : REAL;
    loLevel : REAL;
    hystWindow : REAL;
END_VAR
VAR_OUTPUT
    hiAlarm : BOOL;
    loAlarm : BOOL;
    error : BOOL;
    status : WORD;
END_VAR
VAR
END_VAR

(* ENGINEERING_CONTRACT
   hiAlarm: retained latch. Activation when Value > hiLevel (PUB001/PUB004).
   Hold until Value < hiLevel - hystWindow (PUB001/PUB004). No external reset.
   loAlarm: retained latch. Activation when Value < loLevel (PUB002/PUB005).
   Hold until Value > loLevel + hystWindow (PUB002/PUB005). No external reset.
   error/status: scan-combinational. Priority loLevel >= hiLevel ->
   error=TRUE, status=16#8001, RETURN (PUB003/PUB006). Else
   hystWindow >= hiLevel - loLevel -> error=TRUE, status=16#8002, RETURN
   (PUB003/PUB007). Else error=FALSE, status=16#0000.
   Error paths exit before alarm evaluation; latched alarm outputs retain
   last values. Unspecified error alarm reset behavior kept as retention.
   Boundaries are strict as stated. *)
(* CONTRACT_RULES [] *)

IF loLevel >= hiLevel THEN
    error := TRUE;
    status := WORD#16#8001;
    RETURN;
END_IF;

IF hystWindow >= (hiLevel - loLevel) THEN
    error := TRUE;
    status := WORD#16#8002;
    RETURN;
END_IF;

error := FALSE;
status := WORD#16#0000;

IF hiAlarm THEN
    IF Value < (hiLevel - hystWindow) THEN
        hiAlarm := FALSE;
    END_IF;
ELSE
    IF Value > hiLevel THEN
        hiAlarm := TRUE;
    END_IF;
END_IF;

IF loAlarm THEN
    IF Value > (loLevel + hystWindow) THEN
        loAlarm := FALSE;
    END_IF;
ELSE
    IF Value < loLevel THEN
        loAlarm := TRUE;
    END_IF;
END_IF;

(* ---- public-easy-03.candidate_02.st ---- *)
FUNCTION_BLOCK AlarmHandling
VAR_INPUT
    Value : REAL;
    hiLevel : REAL;
    loLevel : REAL;
    hystWindow : REAL;
END_VAR
VAR_OUTPUT
    hiAlarm : BOOL;
    loAlarm : BOOL;
    error : BOOL;
    status : WORD;
END_VAR
VAR
END_VAR

(* ENGINEERING_CONTRACT
   hiAlarm: retained latch. Activation when Value > hiLevel (PUB001/PUB004).
   Hold until Value < hiLevel - hystWindow (PUB001/PUB004). No external reset.
   loAlarm: retained latch. Activation when Value < loLevel (PUB002/PUB005).
   Hold until Value > loLevel + hystWindow (PUB002/PUB005). No external reset.
   error/status: scan-combinational. Priority loLevel >= hiLevel ->
   error=TRUE, status=16#8001, RETURN (PUB003/PUB006). Else
   hystWindow >= hiLevel - loLevel -> error=TRUE, status=16#8002, RETURN
   (PUB003/PUB007). Else error=FALSE, status=16#0000.
   Error paths exit before alarm evaluation; latched alarm outputs retain
   last values. Unspecified error alarm reset behavior kept as retention.
   Boundaries are strict as stated. *)
(* CONTRACT_RULES [] *)

IF loLevel >= hiLevel THEN
    error := TRUE;
    status := WORD#16#8001;
    RETURN;
END_IF;

IF hystWindow >= (hiLevel - loLevel) THEN
    error := TRUE;
    status := WORD#16#8002;
    RETURN;
END_IF;

error := FALSE;
status := WORD#16#0000;

IF hiAlarm THEN
    IF Value < (hiLevel - hystWindow) THEN
        hiAlarm := FALSE;
    END_IF;
ELSE
    IF Value > hiLevel THEN
        hiAlarm := TRUE;
    END_IF;
END_IF;

IF loAlarm THEN
    IF Value > (loLevel + hystWindow) THEN
        loAlarm := FALSE;
    END_IF;
ELSE
    IF Value < loLevel THEN
        loAlarm := TRUE;
    END_IF;
END_IF;

END_FUNCTION_BLOCK

(* ---- public-easy-03.raw_candidate_01.st ---- *)
FUNCTION_BLOCK AlarmHandling
VAR_INPUT
    Value : REAL;
    hiLevel : REAL;
    loLevel : REAL;
    hystWindow : REAL;
END_VAR
VAR_OUTPUT
    hiAlarm : BOOL;
    loAlarm : BOOL;
    error : BOOL;
    status : WORD;
END_VAR
VAR
END_VAR

(* ENGINEERING_CONTRACT
   hiAlarm: retained latch. Activation when Value > hiLevel (PUB001/PUB004).
   Hold until Value < hiLevel - hystWindow (PUB001/PUB004). No external reset.
   loAlarm: retained latch. Activation when Value < loLevel (PUB002/PUB005).
   Hold until Value > loLevel + hystWindow (PUB002/PUB005). No external reset.
   error/status: scan-combinational. Priority loLevel >= hiLevel ->
   error=TRUE, status=16#8001, RETURN (PUB003/PUB006). Else
   hystWindow >= hiLevel - loLevel -> error=TRUE, status=16#8002, RETURN
   (PUB003/PUB007). Else error=FALSE, status=16#0000.
   Error paths exit before alarm evaluation; latched alarm outputs retain
   last values. Unspecified error alarm reset behavior kept as retention.
   Boundaries are strict as stated. *)
(* CONTRACT_RULES [] *)

IF loLevel >= hiLevel THEN
    error := TRUE;
    status := WORD#16#8001;
    RETURN;
END_IF;

IF hystWindow >= (hiLevel - loLevel) THEN
    error := TRUE;
    status := WORD#16#8002;
    RETURN;
END_IF;

error := FALSE;
status := WORD#16#0000;

IF hiAlarm THEN
    IF Value < (hiLevel - hystWindow) THEN
        hiAlarm := FALSE;
    END_IF;
ELSE
    IF Value > hiLevel THEN
        hiAlarm := TRUE;
    END_IF;
END_IF;

IF loAlarm THEN
    IF Value > (loLevel + hystWindow) THEN
        loAlarm := FALSE;
    END_IF;
ELSE
    IF Value < loLevel THEN
        loAlarm := TRUE;
    END_IF;
END_IF;

(* ---- public-easy-03.raw_candidate_02.st ---- *)
FUNCTION_BLOCK AlarmHandling
VAR_INPUT
    Value : REAL;
    hiLevel : REAL;
    loLevel : REAL;
    hystWindow : REAL;
END_VAR
VAR_OUTPUT
    hiAlarm : BOOL;
    loAlarm : BOOL;
    error : BOOL;
    status : WORD;
END_VAR
VAR
END_VAR

(* ENGINEERING_CONTRACT
   hiAlarm: retained latch. Activation when Value > hiLevel (PUB001/PUB004).
   Hold until Value < hiLevel - hystWindow (PUB001/PUB004). No external reset.
   loAlarm: retained latch. Activation when Value < loLevel (PUB002/PUB005).
   Hold until Value > loLevel + hystWindow (PUB002/PUB005). No external reset.
   error/status: scan-combinational. Priority loLevel >= hiLevel ->
   error=TRUE, status=16#8001, RETURN (PUB003/PUB006). Else
   hystWindow >= hiLevel - loLevel -> error=TRUE, status=16#8002, RETURN
   (PUB003/PUB007). Else error=FALSE, status=16#0000.
   Error paths exit before alarm evaluation; latched alarm outputs retain
   last values. Unspecified error alarm reset behavior kept as retention.
   Boundaries are strict as stated. *)
(* CONTRACT_RULES [] *)

IF loLevel >= hiLevel THEN
    error := TRUE;
    status := WORD#16#8001;
    RETURN;
END_IF;

IF hystWindow >= (hiLevel - loLevel) THEN
    error := TRUE;
    status := WORD#16#8002;
    RETURN;
END_IF;

error := FALSE;
status := WORD#16#0000;

IF hiAlarm THEN
    IF Value < (hiLevel - hystWindow) THEN
        hiAlarm := FALSE;
    END_IF;
ELSE
    IF Value > hiLevel THEN
        hiAlarm := TRUE;
    END_IF;
END_IF;

IF loAlarm THEN
    IF Value > (loLevel + hystWindow) THEN
        loAlarm := FALSE;
    END_IF;
ELSE
    IF Value < loLevel THEN
        loAlarm := TRUE;
    END_IF;
END_IF;

END_FUNCTION_BLOCK

(* ---- public-easy-04.candidate_01.st ---- *)
(*
ENGINEERING_CONTRACT
- VFD_RUN: combinational; TRUE only when PASTE_E_STOP_NC TRUE and debounced viscosity valid; no retention; E-stop FALSE immediately disables (PUB002).
- Viscosity debounce: TON IN = VISCOSITY_OK AND NOT(incomplete AND E-stop FALSE); VISCOSITY_OK FALSE invalidates immediately; E-stop clears incomplete debounce only (PUB001,PUB002).
- Accumulator: updates by TO_LTIME(CycleTime) only while VFD_RUN TRUE this scan; otherwise holds; initial LTIME#0s (PUB003,PUB005).
- Maintenance: computed as accumulated >= LTIME#500h, informational only, remains TRUE while runtime above threshold, no reset (PUB004).
- Units: DebounceTime/CycleTime are TIME; runtime/output are LTIME; threshold uses >= boundary (PUB004).
*)
(* CONTRACT_RULES [] *)
FUNCTION_BLOCK FB_JamPumpDebouncingRuntime
VAR_INPUT
    VISCOSITY_OK : BOOL;
    PASTE_E_STOP_NC : BOOL;
    DebounceTime : TIME;
    CycleTime : TIME;
END_VAR
VAR_OUTPUT
    VFD_RUN : BOOL := FALSE;
    PUMP_MAINT_DUE : BOOL := FALSE;
    PUMP_RUNTIME_ACC : LTIME := LTIME#0s;
END_VAR
VAR
    tmp_DebounceTimer : TON;
    tmp_PrevDebounceQ : BOOL;
    tmp_EStopClearIncomplete : BOOL;
    tmp_Debounced : BOOL;
    tmp_RuntimeAcc : LTIME := LTIME#0s;
    tmp_MaintenanceLimit : LTIME := LTIME#500h;
END_VAR

tmp_PrevDebounceQ := tmp_DebounceTimer.Q;
tmp_EStopClearIncomplete := (NOT PASTE_E_STOP_NC) AND (NOT tmp_PrevDebounceQ);

tmp_DebounceTimer(IN := VISCOSITY_OK AND (NOT tmp_EStopClearIncomplete),
                 PT := DebounceTime);
tmp_Debounced := tmp_DebounceTimer.Q;

VFD_RUN := PASTE_E_STOP_NC AND tmp_Debounced;

IF VFD_RUN THEN
    tmp_RuntimeAcc := tmp_RuntimeAcc + TO_LTIME(CycleTime);
END_IF;

PUMP_RUNTIME_ACC := tmp_RuntimeAcc;
PUMP_MAINT_DUE := (tmp_RuntimeAcc >= tmp_MaintenanceLimit);

(* ---- public-easy-04.candidate_02.st ---- *)
(*
ENGINEERING_CONTRACT
- VFD_RUN: combinational; TRUE only when PASTE_E_STOP_NC TRUE and debounced viscosity valid; no retention; E-stop FALSE immediately disables (PUB002).
- Viscosity debounce: TON IN = VISCOSITY_OK AND NOT(incomplete AND E-stop FALSE); VISCOSITY_OK FALSE invalidates immediately; E-stop clears incomplete debounce only (PUB001,PUB002).
- Accumulator: updates by TO_LTIME(CycleTime) only while VFD_RUN TRUE this scan; otherwise holds; initial LTIME#0s (PUB003,PUB005).
- Maintenance: computed as accumulated >= LTIME#500h, informational only, remains TRUE while runtime above threshold, no reset (PUB004).
- Units: DebounceTime/CycleTime are TIME; runtime/output are LTIME; threshold uses >= boundary (PUB004).
*)
(* CONTRACT_RULES [] *)
FUNCTION_BLOCK FB_JamPumpDebouncingRuntime
VAR_INPUT
    VISCOSITY_OK : BOOL;
    PASTE_E_STOP_NC : BOOL;
    DebounceTime : TIME;
    CycleTime : TIME;
END_VAR
VAR_OUTPUT
    VFD_RUN : BOOL := FALSE;
    PUMP_MAINT_DUE : BOOL := FALSE;
    PUMP_RUNTIME_ACC : LTIME := LTIME#0s;
END_VAR
VAR
    tmp_DebounceTimer : TON;
    tmp_PrevDebounceQ : BOOL;
    tmp_EStopClearIncomplete : BOOL;
    tmp_Debounced : BOOL;
    tmp_RuntimeAcc : LTIME := LTIME#0s;
    tmp_MaintenanceLimit : LTIME := LTIME#500h;
END_VAR

tmp_PrevDebounceQ := tmp_DebounceTimer.Q;
tmp_EStopClearIncomplete := (NOT PASTE_E_STOP_NC) AND (NOT tmp_PrevDebounceQ);

tmp_DebounceTimer(IN := VISCOSITY_OK AND (NOT tmp_EStopClearIncomplete),
                 PT := DebounceTime);
tmp_Debounced := tmp_DebounceTimer.Q;

VFD_RUN := PASTE_E_STOP_NC AND tmp_Debounced;

IF VFD_RUN THEN
    tmp_RuntimeAcc := tmp_RuntimeAcc + TO_LTIME(CycleTime);
END_IF;

PUMP_RUNTIME_ACC := tmp_RuntimeAcc;
PUMP_MAINT_DUE := (tmp_RuntimeAcc >= tmp_MaintenanceLimit);

END_FUNCTION_BLOCK

(* ---- public-easy-04.raw_candidate_01.st ---- *)
(*
ENGINEERING_CONTRACT
- VFD_RUN: combinational; TRUE only when PASTE_E_STOP_NC TRUE and debounced viscosity valid; no retention; E-stop FALSE immediately disables (PUB002).
- Viscosity debounce: TON IN = VISCOSITY_OK AND NOT(incomplete AND E-stop FALSE); VISCOSITY_OK FALSE invalidates immediately; E-stop clears incomplete debounce only (PUB001,PUB002).
- Accumulator: updates by TO_LTIME(CycleTime) only while VFD_RUN TRUE this scan; otherwise holds; initial LTIME#0s (PUB003,PUB005).
- Maintenance: computed as accumulated >= LTIME#500h, informational only, remains TRUE while runtime above threshold, no reset (PUB004).
- Units: DebounceTime/CycleTime are TIME; runtime/output are LTIME; threshold uses >= boundary (PUB004).
*)
(* CONTRACT_RULES [] *)
FUNCTION_BLOCK FB_JamPumpDebouncingRuntime
VAR_INPUT
    VISCOSITY_OK : BOOL;
    PASTE_E_STOP_NC : BOOL;
    DebounceTime : TIME;
    CycleTime : TIME;
END_VAR
VAR_OUTPUT
    VFD_RUN : BOOL := FALSE;
    PUMP_MAINT_DUE : BOOL := FALSE;
    PUMP_RUNTIME_ACC : LTIME := LTIME#0s;
END_VAR
VAR
    tmp_DebounceTimer : TON;
    tmp_PrevDebounceQ : BOOL;
    tmp_EStopClearIncomplete : BOOL;
    tmp_Debounced : BOOL;
    tmp_RuntimeAcc : LTIME := LTIME#0s;
    tmp_MaintenanceLimit : LTIME := LTIME#500h;
END_VAR

tmp_PrevDebounceQ := tmp_DebounceTimer.Q;
tmp_EStopClearIncomplete := (NOT PASTE_E_STOP_NC) AND (NOT tmp_PrevDebounceQ);

tmp_DebounceTimer(IN := VISCOSITY_OK AND (NOT tmp_EStopClearIncomplete),
                 PT := DebounceTime);
tmp_Debounced := tmp_DebounceTimer.Q;

VFD_RUN := PASTE_E_STOP_NC AND tmp_Debounced;

IF VFD_RUN THEN
    tmp_RuntimeAcc := tmp_RuntimeAcc + TO_LTIME(CycleTime);
END_IF;

PUMP_RUNTIME_ACC := tmp_RuntimeAcc;
PUMP_MAINT_DUE := (tmp_RuntimeAcc >= tmp_MaintenanceLimit);

(* ---- public-easy-04.raw_candidate_02.st ---- *)
(*
ENGINEERING_CONTRACT
- VFD_RUN: combinational; TRUE only when PASTE_E_STOP_NC TRUE and debounced viscosity valid; no retention; E-stop FALSE immediately disables (PUB002).
- Viscosity debounce: TON IN = VISCOSITY_OK AND NOT(incomplete AND E-stop FALSE); VISCOSITY_OK FALSE invalidates immediately; E-stop clears incomplete debounce only (PUB001,PUB002).
- Accumulator: updates by TO_LTIME(CycleTime) only while VFD_RUN TRUE this scan; otherwise holds; initial LTIME#0s (PUB003,PUB005).
- Maintenance: computed as accumulated >= LTIME#500h, informational only, remains TRUE while runtime above threshold, no reset (PUB004).
- Units: DebounceTime/CycleTime are TIME; runtime/output are LTIME; threshold uses >= boundary (PUB004).
*)
(* CONTRACT_RULES [] *)
FUNCTION_BLOCK FB_JamPumpDebouncingRuntime
VAR_INPUT
    VISCOSITY_OK : BOOL;
    PASTE_E_STOP_NC : BOOL;
    DebounceTime : TIME;
    CycleTime : TIME;
END_VAR
VAR_OUTPUT
    VFD_RUN : BOOL := FALSE;
    PUMP_MAINT_DUE : BOOL := FALSE;
    PUMP_RUNTIME_ACC : LTIME := LTIME#0s;
END_VAR
VAR
    tmp_DebounceTimer : TON;
    tmp_PrevDebounceQ : BOOL;
    tmp_EStopClearIncomplete : BOOL;
    tmp_Debounced : BOOL;
    tmp_RuntimeAcc : LTIME := LTIME#0s;
    tmp_MaintenanceLimit : LTIME := LTIME#500h;
END_VAR

tmp_PrevDebounceQ := tmp_DebounceTimer.Q;
tmp_EStopClearIncomplete := (NOT PASTE_E_STOP_NC) AND (NOT tmp_PrevDebounceQ);

tmp_DebounceTimer(IN := VISCOSITY_OK AND (NOT tmp_EStopClearIncomplete),
                 PT := DebounceTime);
tmp_Debounced := tmp_DebounceTimer.Q;

VFD_RUN := PASTE_E_STOP_NC AND tmp_Debounced;

IF VFD_RUN THEN
    tmp_RuntimeAcc := tmp_RuntimeAcc + TO_LTIME(CycleTime);
END_IF;

PUMP_RUNTIME_ACC := tmp_RuntimeAcc;
PUMP_MAINT_DUE := (tmp_RuntimeAcc >= tmp_MaintenanceLimit);

END_FUNCTION_BLOCK

(* ---- public-easy-05.candidate_01.st ---- *)
FUNCTION_BLOCK WeldGapAlarm
VAR_INPUT
    Gap_Exceeded : BOOL;
    Weld_E_Stop_NC : BOOL;
    DebounceTime : TIME;
END_VAR
VAR_OUTPUT
    Operator_Alert : BOOL;
    Weld_Soft_Start_Active : BOOL;
END_VAR
VAR
    InitTimer : TON;
    DebounceTimer : TON;
END_VAR

(* ENGINEERING_CONTRACT
Operator_Alert:
  activation: InitTimer.Q AND Weld_E_Stop_NC AND DebounceTimer.Q (PUB003/PUB004)
  hold: remains TRUE only while activation condition is true each scan; no separate latch
  reset/deactivation: Gap_Exceeded FALSE, Weld_E_Stop_NC FALSE, or initialization active
  priority: E-Stop FALSE immediately clears debounce and output; initialization also forces FALSE
  units/boundary: BOOL; DebounceTime is TIME, alert only after Gap_Exceeded remains TRUE >= DebounceTime

Weld_Soft_Start_Active:
  activation: NOT InitTimer.Q, i.e. during first 5 s after power-up (PUB002/PUB005)
  hold: remains TRUE for the entire 5 s initialization window
  reset/deactivation: InitTimer.Q becomes TRUE at >= 5 s
  priority: E-Stop does not deassert this output; PUB004 omits it, so timer status is preserved
  units/boundary: BOOL; 5 s inclusive at timer Q edge

InitTimer:
  unconditional TON with PT := T#5S from first scan; Q is FALSE until ET >= 5 s, then TRUE
DebounceTimer:
  accumulates only when InitTimer.Q AND Weld_E_Stop_NC AND Gap_Exceeded
  reset: Gap_Exceeded FALSE, Weld_E_Stop_NC FALSE, or initialization active
  units: TIME; positive DebounceTime assumed per interface
*)

InitTimer(IN := TRUE, PT := T#5S);

DebounceTimer(
    IN := InitTimer.Q AND Weld_E_Stop_NC AND Gap_Exceeded,
    PT := DebounceTime
);

Weld_Soft_Start_Active := NOT InitTimer.Q;
Operator_Alert := Weld_E_Stop_NC AND DebounceTimer.Q;

(* CONTRACT_RULES [] *)

END_FUNCTION_BLOCK

(* ---- public-easy-05.raw_candidate_01.st ---- *)
FUNCTION_BLOCK WeldGapAlarm
VAR_INPUT
    Gap_Exceeded : BOOL;
    Weld_E_Stop_NC : BOOL;
    DebounceTime : TIME;
END_VAR
VAR_OUTPUT
    Operator_Alert : BOOL;
    Weld_Soft_Start_Active : BOOL;
END_VAR
VAR
    InitTimer : TON;
    DebounceTimer : TON;
END_VAR

(* ENGINEERING_CONTRACT
Operator_Alert:
  activation: InitTimer.Q AND Weld_E_Stop_NC AND DebounceTimer.Q (PUB003/PUB004)
  hold: remains TRUE only while activation condition is true each scan; no separate latch
  reset/deactivation: Gap_Exceeded FALSE, Weld_E_Stop_NC FALSE, or initialization active
  priority: E-Stop FALSE immediately clears debounce and output; initialization also forces FALSE
  units/boundary: BOOL; DebounceTime is TIME, alert only after Gap_Exceeded remains TRUE >= DebounceTime

Weld_Soft_Start_Active:
  activation: NOT InitTimer.Q, i.e. during first 5 s after power-up (PUB002/PUB005)
  hold: remains TRUE for the entire 5 s initialization window
  reset/deactivation: InitTimer.Q becomes TRUE at >= 5 s
  priority: E-Stop does not deassert this output; PUB004 omits it, so timer status is preserved
  units/boundary: BOOL; 5 s inclusive at timer Q edge

InitTimer:
  unconditional TON with PT := T#5S from first scan; Q is FALSE until ET >= 5 s, then TRUE
DebounceTimer:
  accumulates only when InitTimer.Q AND Weld_E_Stop_NC AND Gap_Exceeded
  reset: Gap_Exceeded FALSE, Weld_E_Stop_NC FALSE, or initialization active
  units: TIME; positive DebounceTime assumed per interface
*)

InitTimer(IN := TRUE, PT := T#5S);

DebounceTimer(
    IN := InitTimer.Q AND Weld_E_Stop_NC AND Gap_Exceeded,
    PT := DebounceTime
);

Weld_Soft_Start_Active := NOT InitTimer.Q;
Operator_Alert := Weld_E_Stop_NC AND DebounceTimer.Q;

(* CONTRACT_RULES [] *)

END_FUNCTION_BLOCK

(* ---- public-easy-06.candidate_01.st ---- *)
FUNCTION_BLOCK AerationBlowerDelayedStart
VAR_INPUT
    DO_LOW : BOOL;
    AERATION_E_STOP_NC : BOOL;
END_VAR
VAR_OUTPUT
    BLOWER_RUN : BOOL := FALSE;
    AERATION_BLOWER_CYCLE_COUNT : UINT := 0;
END_VAR
VAR
    local_startTimer : TON;
    local_runRise : R_TRIG;
END_VAR

(* ENGINEERING_CONTRACT
BLOWER_RUN:
  Activation: TON.Q becomes TRUE when DO_LOW AND AERATION_E_STOP_NC have remained TRUE for >= 5 s (PUB001).
  Retention/hold: remains TRUE while TON.Q stays TRUE with both input conditions TRUE (PUB001).
  Explicit reset/deactivation: immediately FALSE when DO_LOW is FALSE or emergency stop active (TON.IN := FALSE) (PUB002).
  Same-scan priority: disable/reset has priority over enable because TON.IN is evaluated first (PUB002).
  Units/boundaries: BOOL, unitless.

AERATION_BLOWER_CYCLE_COUNT:
  Activation/update: increments once on a FALSE-to-TRUE transition of BLOWER_RUN, detected by R_TRIG (PUB003).
  Retention/hold: retained between scans; no explicit reset specified (PUB003).
  Same-scan priority: updated after BLOWER_RUN is computed in the same scan (PUB003).
  Units/boundaries: UINT start count, initialized to 0; standard UINT wrap behavior at 65535 (PUB004).
*)

(* CONTRACT_RULES [] *)

local_startTimer(IN := DO_LOW AND AERATION_E_STOP_NC, PT := T#5S);
BLOWER_RUN := local_startTimer.Q;
local_runRise(CLK := BLOWER_RUN);
IF local_runRise.Q THEN
    AERATION_BLOWER_CYCLE_COUNT := AERATION_BLOWER_CYCLE_COUNT + UINT#1;
END_IF;

END_FUNCTION_BLOCK

(* ---- public-easy-06.raw_candidate_01.st ---- *)
FUNCTION_BLOCK AerationBlowerDelayedStart
VAR_INPUT
    DO_LOW : BOOL;
    AERATION_E_STOP_NC : BOOL;
END_VAR
VAR_OUTPUT
    BLOWER_RUN : BOOL := FALSE;
    AERATION_BLOWER_CYCLE_COUNT : UINT := 0;
END_VAR
VAR
    local_startTimer : TON;
    local_runRise : R_TRIG;
END_VAR

(* ENGINEERING_CONTRACT
BLOWER_RUN:
  Activation: TON.Q becomes TRUE when DO_LOW AND AERATION_E_STOP_NC have remained TRUE for >= 5 s (PUB001).
  Retention/hold: remains TRUE while TON.Q stays TRUE with both input conditions TRUE (PUB001).
  Explicit reset/deactivation: immediately FALSE when DO_LOW is FALSE or emergency stop active (TON.IN := FALSE) (PUB002).
  Same-scan priority: disable/reset has priority over enable because TON.IN is evaluated first (PUB002).
  Units/boundaries: BOOL, unitless.

AERATION_BLOWER_CYCLE_COUNT:
  Activation/update: increments once on a FALSE-to-TRUE transition of BLOWER_RUN, detected by R_TRIG (PUB003).
  Retention/hold: retained between scans; no explicit reset specified (PUB003).
  Same-scan priority: updated after BLOWER_RUN is computed in the same scan (PUB003).
  Units/boundaries: UINT start count, initialized to 0; standard UINT wrap behavior at 65535 (PUB004).
*)

(* CONTRACT_RULES [] *)

local_startTimer(IN := DO_LOW AND AERATION_E_STOP_NC, PT := T#5S);
BLOWER_RUN := local_startTimer.Q;
local_runRise(CLK := BLOWER_RUN);
IF local_runRise.Q THEN
    AERATION_BLOWER_CYCLE_COUNT := AERATION_BLOWER_CYCLE_COUNT + UINT#1;
END_IF;

END_FUNCTION_BLOCK

(* ---- public-hard-01.candidate_01.st ---- *)
TYPE AutoState : (ST_IDLE, ST_OPEN_A, ST_OPEN_B, ST_OPEN_C, ST_MIXING);
END_TYPE;

FUNCTION_BLOCK MaterialProportioningControl
VAR_INPUT
    estop : BOOL;
    opeMode : BOOL;
    valveAStart : BOOL;
    valveBStart : BOOL;
    valveCStart : BOOL;
    valveDStart : BOOL;
    mixMotorStart : BOOL;
    autoStart : BOOL;
    processMode : BOOL;
    levelSensor : INT;
    mixMotorComplete : BOOL;
END_VAR
VAR_OUTPUT
    valveARun : BOOL;
    valveBRun : BOOL;
    valveCRun : BOOL;
    valveDRun : BOOL;
    mixMotorRun : BOOL;
END_VAR
VAR
    trigA : R_TRIG;
    trigB : R_TRIG;
    trigC : R_TRIG;
    trigD : R_TRIG;
    trigMix : R_TRIG;
    trigAuto : R_TRIG;

    manualA : BOOL := FALSE;
    manualB : BOOL := FALSE;
    manualC : BOOL := FALSE;
    manualD : BOOL := FALSE;
    manualMixer : BOOL := FALSE;

    autoActive : BOOL := FALSE;
    autoState : AutoState := ST_IDLE;
    finalDCommand : BOOL := FALSE;
END_VAR

(* ENGINEERING_CONTRACT
Manual outputs: set/toggled on rising edge of each start input while opeMode=FALSE.
Manual outputs retain until next rising edge of same input or estop=FALSE.
Automatic sequence outputs: activated by autoStart rising edge while opeMode=TRUE and not already active.
State thresholds: levelSensor >= 50 (A->B), >= 80 (B->C or B->mix), >= 100 (C->mix).
processMode is evaluated at the 80 cm transition only.
Mixer stops and valve D opens on mixMotorComplete=TRUE while mixing.
valveDRun remains held by finalDCommand after automatic process ends until next autoStart or estop.
Priority: estop=FALSE forces all outputs FALSE and resets all manual/automatic state.
Same-scan: autoStart sets ST_OPEN_A and outputs without immediate threshold transition; other transitions are one state per scan.
Units: levelSensor cm. PUB001-PUB015.
*)

(* CONTRACT_RULES [] *)

// Rising-edge detection is updated every scan, including during emergency stop.
trigA(CLK := valveAStart);
trigB(CLK := valveBStart);
trigC(CLK := valveCStart);
trigD(CLK := valveDStart);
trigMix(CLK := mixMotorStart);
trigAuto(CLK := autoStart);

IF NOT estop THEN
    // Emergency stop: stop everything immediately and reset all retained state.
    valveARun := FALSE;
    valveBRun := FALSE;
    valveCRun := FALSE;
    valveDRun := FALSE;
    mixMotorRun := FALSE;

    manualA := FALSE;
    manualB := FALSE;
    manualC := FALSE;
    manualD := FALSE;
    manualMixer := FALSE;

    autoActive := FALSE;
    autoState := ST_IDLE;
    finalDCommand := FALSE;

    RETURN;
END_IF;

IF NOT opeMode THEN
    // Manual operation mode.
    IF trigA.Q THEN
        manualA := NOT manualA;
    END_IF;
    IF trigB.Q THEN
        manualB := NOT manualB;
    END_IF;
    IF trigC.Q THEN
        manualC := NOT manualC;
    END_IF;
    IF trigD.Q THEN
        manualD := NOT manualD;
    END_IF;
    IF trigMix.Q THEN
        manualMixer := NOT manualMixer;
    END_IF;

    valveARun := manualA;
    valveBRun := manualB;
    valveCRun := manualC;
    valveDRun := manualD;
    mixMotorRun := manualMixer;

ELSE
    // Automatic operation mode.
    IF trigAuto.Q AND NOT autoActive THEN
        // Start new automatic process: open valve A first.
        autoActive := TRUE;
        autoState := ST_OPEN_A;
        finalDCommand := FALSE;

        valveARun := TRUE;
        valveBRun := FALSE;
        valveCRun := FALSE;
        valveDRun := FALSE;
        mixMotorRun := FALSE;
    ELSE
        CASE autoState OF
            ST_IDLE:
                valveARun := FALSE;
                valveBRun := FALSE;
                valveCRun := FALSE;
                valveDRun := finalDCommand;
                mixMotorRun := FALSE;

            ST_OPEN_A:
                valveARun := TRUE;
                valveBRun := FALSE;
                valveCRun := FALSE;
                valveDRun := FALSE;
                mixMotorRun := FALSE;

                IF levelSensor >= 50 THEN
                    autoState := ST_OPEN_B;
                    valveARun := FALSE;
                    valveBRun := TRUE;
                END_IF;

            ST_OPEN_B:
                valveARun := FALSE;
                valveBRun := TRUE;
                valveCRun := FALSE;
                valveDRun := FALSE;
                mixMotorRun := FALSE;

                IF levelSensor >= 80 THEN
                    IF NOT processMode THEN
                        // processMode = FALSE: close B, start mixer.
                        autoState := ST_MIXING;
                        valveBRun := FALSE;
                        mixMotorRun := TRUE;
                    ELSE
                        // processMode = TRUE: close B, open C.
                        autoState := ST_OPEN_C;
                        valveBRun := FALSE;
                        valveCRun := TRUE;
                    END_IF;
                END_IF;

            ST_OPEN_C:
                valveARun := FALSE;
                valveBRun := FALSE;
                valveCRun := TRUE;
                valveDRun := FALSE;
                mixMotorRun := FALSE;

                IF levelSensor >= 100 THEN
                    autoState := ST_MIXING;
                    valveCRun := FALSE;
                    mixMotorRun := TRUE;
                END_IF;

            ST_MIXING:
                valveARun := FALSE;
                valveBRun := FALSE;
                valveCRun := FALSE;
                valveDRun := FALSE;
                mixMotorRun := TRUE;

                IF mixMotorComplete THEN
                    mixMotorRun := FALSE;
                    valveDRun := TRUE;
                    finalDCommand := TRUE;
                    autoActive := FALSE;
                    autoState := ST_IDLE;
                END_IF;
        END_CASE;
    END_IF;
END_IF;

(* ---- public-hard-01.candidate_02.st ---- *)
TYPE AutoState : (ST_IDLE, ST_OPEN_A, ST_OPEN_B, ST_OPEN_C, ST_MIXING);
END_TYPE;

FUNCTION_BLOCK MaterialProportioningControl
VAR_INPUT
    estop : BOOL;
    opeMode : BOOL;
    valveAStart : BOOL;
    valveBStart : BOOL;
    valveCStart : BOOL;
    valveDStart : BOOL;
    mixMotorStart : BOOL;
    autoStart : BOOL;
    processMode : BOOL;
    levelSensor : INT;
    mixMotorComplete : BOOL;
END_VAR
VAR_OUTPUT
    valveARun : BOOL;
    valveBRun : BOOL;
    valveCRun : BOOL;
    valveDRun : BOOL;
    mixMotorRun : BOOL;
END_VAR
VAR
    trigA : R_TRIG;
    trigB : R_TRIG;
    trigC : R_TRIG;
    trigD : R_TRIG;
    trigMix : R_TRIG;
    trigAuto : R_TRIG;

    manualA : BOOL := FALSE;
    manualB : BOOL := FALSE;
    manualC : BOOL := FALSE;
    manualD : BOOL := FALSE;
    manualMixer : BOOL := FALSE;

    autoActive : BOOL := FALSE;
    autoState : AutoState := ST_IDLE;
    finalDCommand : BOOL := FALSE;
END_VAR

(* ENGINEERING_CONTRACT
Manual outputs: set/toggled on rising edge of each start input while opeMode=FALSE.
Manual outputs retain until next rising edge of same input or estop=FALSE.
Automatic sequence outputs: activated by autoStart rising edge while opeMode=TRUE and not already active.
State thresholds: levelSensor >= 50 (A->B), >= 80 (B->C or B->mix), >= 100 (C->mix).
processMode is evaluated at the 80 cm transition only.
Mixer stops and valve D opens on mixMotorComplete=TRUE while mixing.
valveDRun remains held by finalDCommand after automatic process ends until next autoStart or estop.
Priority: estop=FALSE forces all outputs FALSE and resets all manual/automatic state.
Same-scan: autoStart sets ST_OPEN_A and outputs without immediate threshold transition; other transitions are one state per scan.
Units: levelSensor cm. PUB001-PUB015.
*)

(* CONTRACT_RULES [] *)

// Rising-edge detection is updated every scan, including during emergency stop.
trigA(CLK := valveAStart);
trigB(CLK := valveBStart);
trigC(CLK := valveCStart);
trigD(CLK := valveDStart);
trigMix(CLK := mixMotorStart);
trigAuto(CLK := autoStart);

IF NOT estop THEN
    // Emergency stop: stop everything immediately and reset all retained state.
    valveARun := FALSE;
    valveBRun := FALSE;
    valveCRun := FALSE;
    valveDRun := FALSE;
    mixMotorRun := FALSE;

    manualA := FALSE;
    manualB := FALSE;
    manualC := FALSE;
    manualD := FALSE;
    manualMixer := FALSE;

    autoActive := FALSE;
    autoState := ST_IDLE;
    finalDCommand := FALSE;

    RETURN;
END_IF;

IF NOT opeMode THEN
    // Manual operation mode.
    IF trigA.Q THEN
        manualA := NOT manualA;
    END_IF;
    IF trigB.Q THEN
        manualB := NOT manualB;
    END_IF;
    IF trigC.Q THEN
        manualC := NOT manualC;
    END_IF;
    IF trigD.Q THEN
        manualD := NOT manualD;
    END_IF;
    IF trigMix.Q THEN
        manualMixer := NOT manualMixer;
    END_IF;

    valveARun := manualA;
    valveBRun := manualB;
    valveCRun := manualC;
    valveDRun := manualD;
    mixMotorRun := manualMixer;

ELSE
    // Automatic operation mode.
    IF trigAuto.Q AND NOT autoActive THEN
        // Start new automatic process: open valve A first.
        autoActive := TRUE;
        autoState := ST_OPEN_A;
        finalDCommand := FALSE;

        valveARun := TRUE;
        valveBRun := FALSE;
        valveCRun := FALSE;
        valveDRun := FALSE;
        mixMotorRun := FALSE;
    ELSE
        CASE autoState OF
            ST_IDLE:
                valveARun := FALSE;
                valveBRun := FALSE;
                valveCRun := FALSE;
                valveDRun := finalDCommand;
                mixMotorRun := FALSE;

            ST_OPEN_A:
                valveARun := TRUE;
                valveBRun := FALSE;
                valveCRun := FALSE;
                valveDRun := FALSE;
                mixMotorRun := FALSE;

                IF levelSensor >= 50 THEN
                    autoState := ST_OPEN_B;
                    valveARun := FALSE;
                    valveBRun := TRUE;
                END_IF;

            ST_OPEN_B:
                valveARun := FALSE;
                valveBRun := TRUE;
                valveCRun := FALSE;
                valveDRun := FALSE;
                mixMotorRun := FALSE;

                IF levelSensor >= 80 THEN
                    IF NOT processMode THEN
                        // processMode = FALSE: close B, start mixer.
                        autoState := ST_MIXING;
                        valveBRun := FALSE;
                        mixMotorRun := TRUE;
                    ELSE
                        // processMode = TRUE: close B, open C.
                        autoState := ST_OPEN_C;
                        valveBRun := FALSE;
                        valveCRun := TRUE;
                    END_IF;
                END_IF;

            ST_OPEN_C:
                valveARun := FALSE;
                valveBRun := FALSE;
                valveCRun := TRUE;
                valveDRun := FALSE;
                mixMotorRun := FALSE;

                IF levelSensor >= 100 THEN
                    autoState := ST_MIXING;
                    valveCRun := FALSE;
                    mixMotorRun := TRUE;
                END_IF;

            ST_MIXING:
                valveARun := FALSE;
                valveBRun := FALSE;
                valveCRun := FALSE;
                valveDRun := FALSE;
                mixMotorRun := TRUE;

                IF mixMotorComplete THEN
                    mixMotorRun := FALSE;
                    valveDRun := TRUE;
                    finalDCommand := TRUE;
                    autoActive := FALSE;
                    autoState := ST_IDLE;
                END_IF;
        END_CASE;
    END_IF;
END_IF;
END_FUNCTION_BLOCK

(* ---- public-hard-01.raw_candidate_01.st ---- *)
TYPE AutoState : (ST_IDLE, ST_OPEN_A, ST_OPEN_B, ST_OPEN_C, ST_MIXING);
END_TYPE

FUNCTION_BLOCK MaterialProportioningControl
VAR_INPUT
    estop : BOOL;
    opeMode : BOOL;
    valveAStart : BOOL;
    valveBStart : BOOL;
    valveCStart : BOOL;
    valveDStart : BOOL;
    mixMotorStart : BOOL;
    autoStart : BOOL;
    processMode : BOOL;
    levelSensor : INT;
    mixMotorComplete : BOOL;
END_VAR
VAR_OUTPUT
    valveARun : BOOL;
    valveBRun : BOOL;
    valveCRun : BOOL;
    valveDRun : BOOL;
    mixMotorRun : BOOL;
END_VAR
VAR
    trigA : R_TRIG;
    trigB : R_TRIG;
    trigC : R_TRIG;
    trigD : R_TRIG;
    trigMix : R_TRIG;
    trigAuto : R_TRIG;

    manualA : BOOL := FALSE;
    manualB : BOOL := FALSE;
    manualC : BOOL := FALSE;
    manualD : BOOL := FALSE;
    manualMixer : BOOL := FALSE;

    autoActive : BOOL := FALSE;
    autoState : AutoState := ST_IDLE;
    finalDCommand : BOOL := FALSE;
END_VAR

(* ENGINEERING_CONTRACT
Manual outputs: set/toggled on rising edge of each start input while opeMode=FALSE.
Manual outputs retain until next rising edge of same input or estop=FALSE.
Automatic sequence outputs: activated by autoStart rising edge while opeMode=TRUE and not already active.
State thresholds: levelSensor >= 50 (A->B), >= 80 (B->C or B->mix), >= 100 (C->mix).
processMode is evaluated at the 80 cm transition only.
Mixer stops and valve D opens on mixMotorComplete=TRUE while mixing.
valveDRun remains held by finalDCommand after automatic process ends until next autoStart or estop.
Priority: estop=FALSE forces all outputs FALSE and resets all manual/automatic state.
Same-scan: autoStart sets ST_OPEN_A and outputs without immediate threshold transition; other transitions are one state per scan.
Units: levelSensor cm. PUB001-PUB015.
*)

(* CONTRACT_RULES [] *)

// Rising-edge detection is updated every scan, including during emergency stop.
trigA(CLK := valveAStart);
trigB(CLK := valveBStart);
trigC(CLK := valveCStart);
trigD(CLK := valveDStart);
trigMix(CLK := mixMotorStart);
trigAuto(CLK := autoStart);

IF NOT estop THEN
    // Emergency stop: stop everything immediately and reset all retained state.
    valveARun := FALSE;
    valveBRun := FALSE;
    valveCRun := FALSE;
    valveDRun := FALSE;
    mixMotorRun := FALSE;

    manualA := FALSE;
    manualB := FALSE;
    manualC := FALSE;
    manualD := FALSE;
    manualMixer := FALSE;

    autoActive := FALSE;
    autoState := ST_IDLE;
    finalDCommand := FALSE;

    RETURN;
END_IF

IF NOT opeMode THEN
    // Manual operation mode.
    IF trigA.Q THEN
        manualA := NOT manualA;
    END_IF;
    IF trigB.Q THEN
        manualB := NOT manualB;
    END_IF;
    IF trigC.Q THEN
        manualC := NOT manualC;
    END_IF;
    IF trigD.Q THEN
        manualD := NOT manualD;
    END_IF;
    IF trigMix.Q THEN
        manualMixer := NOT manualMixer;
    END_IF;

    valveARun := manualA;
    valveBRun := manualB;
    valveCRun := manualC;
    valveDRun := manualD;
    mixMotorRun := manualMixer;

ELSE
    // Automatic operation mode.
    IF trigAuto.Q AND NOT autoActive THEN
        // Start new automatic process: open valve A first.
        autoActive := TRUE;
        autoState := ST_OPEN_A;
        finalDCommand := FALSE;

        valveARun := TRUE;
        valveBRun := FALSE;
        valveCRun := FALSE;
        valveDRun := FALSE;
        mixMotorRun := FALSE;
    ELSE
        CASE autoState OF
            ST_IDLE:
                valveARun := FALSE;
                valveBRun := FALSE;
                valveCRun := FALSE;
                valveDRun := finalDCommand;
                mixMotorRun := FALSE;

            ST_OPEN_A:
                valveARun := TRUE;
                valveBRun := FALSE;
                valveCRun := FALSE;
                valveDRun := FALSE;
                mixMotorRun := FALSE;

                IF levelSensor >= 50 THEN
                    autoState := ST_OPEN_B;
                    valveARun := FALSE;
                    valveBRun := TRUE;
                END_IF;

            ST_OPEN_B:
                valveARun := FALSE;
                valveBRun := TRUE;
                valveCRun := FALSE;
                valveDRun := FALSE;
                mixMotorRun := FALSE;

                IF levelSensor >= 80 THEN
                    IF NOT processMode THEN
                        // processMode = FALSE: close B, start mixer.
                        autoState := ST_MIXING;
                        valveBRun := FALSE;
                        mixMotorRun := TRUE;
                    ELSE
                        // processMode = TRUE: close B, open C.
                        autoState := ST_OPEN_C;
                        valveBRun := FALSE;
                        valveCRun := TRUE;
                    END_IF;
                END_IF;

            ST_OPEN_C:
                valveARun := FALSE;
                valveBRun := FALSE;
                valveCRun := TRUE;
                valveDRun := FALSE;
                mixMotorRun := FALSE;

                IF levelSensor >= 100 THEN
                    autoState := ST_MIXING;
                    valveCRun := FALSE;
                    mixMotorRun := TRUE;
                END_IF;

            ST_MIXING:
                valveARun := FALSE;
                valveBRun := FALSE;
                valveCRun := FALSE;
                valveDRun := FALSE;
                mixMotorRun := TRUE;

                IF mixMotorComplete THEN
                    mixMotorRun := FALSE;
                    valveDRun := TRUE;
                    finalDCommand := TRUE;
                    autoActive := FALSE;
                    autoState := ST_IDLE;
                END_IF;
        END_CASE;
    END_IF;
END_IF;

(* ---- public-hard-01.raw_candidate_02.st ---- *)
TYPE AutoState : (ST_IDLE, ST_OPEN_A, ST_OPEN_B, ST_OPEN_C, ST_MIXING);
END_TYPE;

FUNCTION_BLOCK MaterialProportioningControl
VAR_INPUT
    estop : BOOL;
    opeMode : BOOL;
    valveAStart : BOOL;
    valveBStart : BOOL;
    valveCStart : BOOL;
    valveDStart : BOOL;
    mixMotorStart : BOOL;
    autoStart : BOOL;
    processMode : BOOL;
    levelSensor : INT;
    mixMotorComplete : BOOL;
END_VAR
VAR_OUTPUT
    valveARun : BOOL;
    valveBRun : BOOL;
    valveCRun : BOOL;
    valveDRun : BOOL;
    mixMotorRun : BOOL;
END_VAR
VAR
    trigA : R_TRIG;
    trigB : R_TRIG;
    trigC : R_TRIG;
    trigD : R_TRIG;
    trigMix : R_TRIG;
    trigAuto : R_TRIG;

    manualA : BOOL := FALSE;
    manualB : BOOL := FALSE;
    manualC : BOOL := FALSE;
    manualD : BOOL := FALSE;
    manualMixer : BOOL := FALSE;

    autoActive : BOOL := FALSE;
    autoState : AutoState := ST_IDLE;
    finalDCommand : BOOL := FALSE;
END_VAR

(* ENGINEERING_CONTRACT
Manual outputs: set/toggled on rising edge of each start input while opeMode=FALSE.
Manual outputs retain until next rising edge of same input or estop=FALSE.
Automatic sequence outputs: activated by autoStart rising edge while opeMode=TRUE and not already active.
State thresholds: levelSensor >= 50 (A->B), >= 80 (B->C or B->mix), >= 100 (C->mix).
processMode is evaluated at the 80 cm transition only.
Mixer stops and valve D opens on mixMotorComplete=TRUE while mixing.
valveDRun remains held by finalDCommand after automatic process ends until next autoStart or estop.
Priority: estop=FALSE forces all outputs FALSE and resets all manual/automatic state.
Same-scan: autoStart sets ST_OPEN_A and outputs without immediate threshold transition; other transitions are one state per scan.
Units: levelSensor cm. PUB001-PUB015.
*)

(* CONTRACT_RULES [] *)

// Rising-edge detection is updated every scan, including during emergency stop.
trigA(CLK := valveAStart);
trigB(CLK := valveBStart);
trigC(CLK := valveCStart);
trigD(CLK := valveDStart);
trigMix(CLK := mixMotorStart);
trigAuto(CLK := autoStart);

IF NOT estop THEN
    // Emergency stop: stop everything immediately and reset all retained state.
    valveARun := FALSE;
    valveBRun := FALSE;
    valveCRun := FALSE;
    valveDRun := FALSE;
    mixMotorRun := FALSE;

    manualA := FALSE;
    manualB := FALSE;
    manualC := FALSE;
    manualD := FALSE;
    manualMixer := FALSE;

    autoActive := FALSE;
    autoState := ST_IDLE;
    finalDCommand := FALSE;

    RETURN;
END_IF;

IF NOT opeMode THEN
    // Manual operation mode.
    IF trigA.Q THEN
        manualA := NOT manualA;
    END_IF;
    IF trigB.Q THEN
        manualB := NOT manualB;
    END_IF;
    IF trigC.Q THEN
        manualC := NOT manualC;
    END_IF;
    IF trigD.Q THEN
        manualD := NOT manualD;
    END_IF;
    IF trigMix.Q THEN
        manualMixer := NOT manualMixer;
    END_IF;

    valveARun := manualA;
    valveBRun := manualB;
    valveCRun := manualC;
    valveDRun := manualD;
    mixMotorRun := manualMixer;

ELSE
    // Automatic operation mode.
    IF trigAuto.Q AND NOT autoActive THEN
        // Start new automatic process: open valve A first.
        autoActive := TRUE;
        autoState := ST_OPEN_A;
        finalDCommand := FALSE;

        valveARun := TRUE;
        valveBRun := FALSE;
        valveCRun := FALSE;
        valveDRun := FALSE;
        mixMotorRun := FALSE;
    ELSE
        CASE autoState OF
            ST_IDLE:
                valveARun := FALSE;
                valveBRun := FALSE;
                valveCRun := FALSE;
                valveDRun := finalDCommand;
                mixMotorRun := FALSE;

            ST_OPEN_A:
                valveARun := TRUE;
                valveBRun := FALSE;
                valveCRun := FALSE;
                valveDRun := FALSE;
                mixMotorRun := FALSE;

                IF levelSensor >= 50 THEN
                    autoState := ST_OPEN_B;
                    valveARun := FALSE;
                    valveBRun := TRUE;
                END_IF;

            ST_OPEN_B:
                valveARun := FALSE;
                valveBRun := TRUE;
                valveCRun := FALSE;
                valveDRun := FALSE;
                mixMotorRun := FALSE;

                IF levelSensor >= 80 THEN
                    IF NOT processMode THEN
                        // processMode = FALSE: close B, start mixer.
                        autoState := ST_MIXING;
                        valveBRun := FALSE;
                        mixMotorRun := TRUE;
                    ELSE
                        // processMode = TRUE: close B, open C.
                        autoState := ST_OPEN_C;
                        valveBRun := FALSE;
                        valveCRun := TRUE;
                    END_IF;
                END_IF;

            ST_OPEN_C:
                valveARun := FALSE;
                valveBRun := FALSE;
                valveCRun := TRUE;
                valveDRun := FALSE;
                mixMotorRun := FALSE;

                IF levelSensor >= 100 THEN
                    autoState := ST_MIXING;
                    valveCRun := FALSE;
                    mixMotorRun := TRUE;
                END_IF;

            ST_MIXING:
                valveARun := FALSE;
                valveBRun := FALSE;
                valveCRun := FALSE;
                valveDRun := FALSE;
                mixMotorRun := TRUE;

                IF mixMotorComplete THEN
                    mixMotorRun := FALSE;
                    valveDRun := TRUE;
                    finalDCommand := TRUE;
                    autoActive := FALSE;
                    autoState := ST_IDLE;
                END_IF;
        END_CASE;
    END_IF;
END_IF;
END_FUNCTION_BLOCK

(* ---- public-hard-02.candidate_01.st ---- *)
TYPE ProcessControl_State : (PC_IDLE, PC_MOVING, PC_WAITING); END_TYPE;

FUNCTION_BLOCK FlexibleProcessingControl
VAR_INPUT
    processLength : USINT;
    sensor1 : BOOL;
    sensor2 : BOOL;
    sensor3 : BOOL;
    sensor4 : BOOL;
    sensor5 : BOOL;
    station1Start : BOOL;
    station2Complete : BOOL;
    station3Complete : BOOL;
    station4Complete : BOOL;
    processSequence : ARRAY[1..8] OF USINT;
END_VAR
VAR_OUTPUT
    conveyorLeft : BOOL;
    conveyorRight : BOOL;
END_VAR
VAR
    state : ProcessControl_State := PC_IDLE;
    currentStation : USINT := 1;
    currentIndex : USINT := 1;
    targetStation : USINT := 0;
    targetSensor : BOOL := FALSE;
    local_rt_start : R_TRIG;
    local_rt_st2 : R_TRIG;
    local_rt_st3 : R_TRIG;
    local_rt_st4 : R_TRIG;
END_VAR

(*
ENGINEERING_CONTRACT
  conveyorLeft / conveyorRight activation: PC_MOVING state and target direction >/< currentStation (PUB001-PUB002).
  Retention/hold: outputs stay on each scan while PC_MOVING until target sensor TRUE (PUB002).
  Explicit reset/deactivation: sensor at target station stops motion and sets both outputs FALSE; next start new product.
  Same-scan priority: start request processed only in PC_IDLE; arrival stop and completion advancement are mutually exclusive by state.
  Units/boundaries: processLength 1..8; processSequence index 1..8; currentStation 1..5; final active entry 5 (PUB003).
  Direction: target > current -> conveyorRight; target < current -> conveyorLeft; target == current -> no movement, treated as arrived.
  Completion edge: rising edge of station2Complete/3/4Complete triggers next step.
  Unspecified: equal consecutive station entries skip movement and wait for completion; simultaneous completion inputs while WAITING use current station only.
*)

(* CONTRACT_RULES [] *)

local_rt_start(CLK := station1Start);
local_rt_st2(CLK := station2Complete);
local_rt_st3(CLK := station3Complete);
local_rt_st4(CLK := station4Complete);

CASE state OF
    PC_IDLE:
        conveyorLeft := FALSE;
        conveyorRight := FALSE;
        IF local_rt_start.Q AND sensor1 THEN
            currentIndex := 1;
            currentStation := 1;
            targetStation := processSequence[currentIndex];
            IF targetStation = currentStation THEN
                IF targetStation = 5 THEN
                    state := PC_IDLE;
                ELSE
                    state := PC_WAITING;
                END_IF;
            ELSE
                state := PC_MOVING;
            END_IF;
        END_IF;

    PC_MOVING:
        targetSensor := FALSE;
        CASE targetStation OF
            2: targetSensor := sensor2;
            3: targetSensor := sensor3;
            4: targetSensor := sensor4;
            5: targetSensor := sensor5;
        END_CASE;

        IF targetStation > currentStation THEN
            conveyorLeft := FALSE;
            conveyorRight := TRUE;
        ELSIF targetStation < currentStation THEN
            conveyorLeft := TRUE;
            conveyorRight := FALSE;
        ELSE
            conveyorLeft := FALSE;
            conveyorRight := FALSE;
        END_IF;

        IF targetSensor THEN
            conveyorLeft := FALSE;
            conveyorRight := FALSE;
            currentStation := targetStation;
            IF targetStation = 5 THEN
                state := PC_IDLE;
            ELSE
                state := PC_WAITING;
            END_IF;
        END_IF;

    PC_WAITING:
        conveyorLeft := FALSE;
        conveyorRight := FALSE;
        IF (currentStation = 2 AND local_rt_st2.Q) OR
           (currentStation = 3 AND local_rt_st3.Q) OR
           (currentStation = 4 AND local_rt_st4.Q) THEN
            IF currentIndex < processLength THEN
                currentIndex := currentIndex + 1;
                targetStation := processSequence[currentIndex];
                IF targetStation = currentStation THEN
                    IF targetStation = 5 THEN
                        state := PC_IDLE;
                    ELSE
                        state := PC_WAITING;
                    END_IF;
                ELSE
                    state := PC_MOVING;
                END_IF;
            ELSE
                state := PC_IDLE;
            END_IF;
        END_IF;
END_CASE;

(* ---- public-hard-02.candidate_02.st ---- *)
TYPE ProcessControl_State : (PC_IDLE, PC_MOVING, PC_WAITING); END_TYPE;

FUNCTION_BLOCK FlexibleProcessingControl
VAR_INPUT
    processLength : USINT;
    sensor1 : BOOL;
    sensor2 : BOOL;
    sensor3 : BOOL;
    sensor4 : BOOL;
    sensor5 : BOOL;
    station1Start : BOOL;
    station2Complete : BOOL;
    station3Complete : BOOL;
    station4Complete : BOOL;
    processSequence : ARRAY[1..8] OF USINT;
END_VAR
VAR_OUTPUT
    conveyorLeft : BOOL;
    conveyorRight : BOOL;
END_VAR
VAR
    state : ProcessControl_State := PC_IDLE;
    currentStation : USINT := 1;
    currentIndex : USINT := 1;
    targetStation : USINT := 0;
    targetSensor : BOOL := FALSE;
    local_rt_start : R_TRIG;
    local_rt_st2 : R_TRIG;
    local_rt_st3 : R_TRIG;
    local_rt_st4 : R_TRIG;
END_VAR

(*
ENGINEERING_CONTRACT
  conveyorLeft / conveyorRight activation: PC_MOVING state and target direction >/< currentStation (PUB001-PUB002).
  Retention/hold: outputs stay on each scan while PC_MOVING until target sensor TRUE (PUB002).
  Explicit reset/deactivation: sensor at target station stops motion and sets both outputs FALSE; next start new product.
  Same-scan priority: start request processed only in PC_IDLE; arrival stop and completion advancement are mutually exclusive by state.
  Units/boundaries: processLength 1..8; processSequence index 1..8; currentStation 1..5; final active entry 5 (PUB003).
  Direction: target > current -> conveyorRight; target < current -> conveyorLeft; target == current -> no movement, treated as arrived.
  Completion edge: rising edge of station2Complete/3/4Complete triggers next step.
  Unspecified: equal consecutive station entries skip movement and wait for completion; simultaneous completion inputs while WAITING use current station only.
*)

(* CONTRACT_RULES [] *)

local_rt_start(CLK := station1Start);
local_rt_st2(CLK := station2Complete);
local_rt_st3(CLK := station3Complete);
local_rt_st4(CLK := station4Complete);

CASE state OF
    PC_IDLE:
        conveyorLeft := FALSE;
        conveyorRight := FALSE;
        IF local_rt_start.Q AND sensor1 THEN
            currentIndex := 1;
            currentStation := 1;
            targetStation := processSequence[currentIndex];
            IF targetStation = currentStation THEN
                IF targetStation = 5 THEN
                    state := PC_IDLE;
                ELSE
                    state := PC_WAITING;
                END_IF;
            ELSE
                state := PC_MOVING;
            END_IF;
        END_IF;

    PC_MOVING:
        targetSensor := FALSE;
        CASE targetStation OF
            2: targetSensor := sensor2;
            3: targetSensor := sensor3;
            4: targetSensor := sensor4;
            5: targetSensor := sensor5;
        END_CASE;

        IF targetStation > currentStation THEN
            conveyorLeft := FALSE;
            conveyorRight := TRUE;
        ELSIF targetStation < currentStation THEN
            conveyorLeft := TRUE;
            conveyorRight := FALSE;
        ELSE
            conveyorLeft := FALSE;
            conveyorRight := FALSE;
        END_IF;

        IF targetSensor THEN
            conveyorLeft := FALSE;
            conveyorRight := FALSE;
            currentStation := targetStation;
            IF targetStation = 5 THEN
                state := PC_IDLE;
            ELSE
                state := PC_WAITING;
            END_IF;
        END_IF;

    PC_WAITING:
        conveyorLeft := FALSE;
        conveyorRight := FALSE;
        IF (currentStation = 2 AND local_rt_st2.Q) OR
           (currentStation = 3 AND local_rt_st3.Q) OR
           (currentStation = 4 AND local_rt_st4.Q) THEN
            IF currentIndex < processLength THEN
                currentIndex := currentIndex + 1;
                targetStation := processSequence[currentIndex];
                IF targetStation = currentStation THEN
                    IF targetStation = 5 THEN
                        state := PC_IDLE;
                    ELSE
                        state := PC_WAITING;
                    END_IF;
                ELSE
                    state := PC_MOVING;
                END_IF;
            ELSE
                state := PC_IDLE;
            END_IF;
        END_IF;
END_CASE;

END_FUNCTION_BLOCK
